(* IEC 61131-3 sources: Industry-PLC-LLM/data/PLCBEAD_repo/PLCBEAD_PLCEmbed-main/PLC-BEAD/Source/PLC_Programs (part 11) *)

(* ---- SIGNAL_4.ST ---- *)
FUNCTION _BYTE_TO_INT:INT
	VAR_INPUT
		IN :	BYTE;
	END_VAR

	_BYTE_TO_INT := USINT_TO_INT(BYTE_TO_USINT(IN));
END_FUNCTION

FUNCTION TIME_TO_UDINT2:UDINT
	VAR_INPUT
		X :	TIME;
	END_VAR

	TIME_TO_UDINT2 := DINT_TO_UDINT(TIME_TO_DINT(X));
END_FUNCTION

FUNCTION UDINT_TO_TIME2:TIME

	VAR_INPUT
		IN :	UDINT;
	END_VAR

	UDINT_TO_TIME2 := DINT_TO_TIME(UDINT_TO_DINT(IN));

END_FUNCTION

FUNCTION_BLOCK T_PLC_MS_block
	VAR_OUTPUT
		T_PLC_MS :	UDINT;
	END_VAR

	VAR_EXTERNAL
		PLC_TICKS_PER_SEC :	INT;
		PLC_SYS_TICK_CNT :	DINT;
	END_VAR

	VAR
		debug :	BOOL;(*Debug-Mode ON / OFF*)
		N :	INT;(*Debug-Faktor*)
		Offset :	UDINT;(*Debug-Offset*)
		temp :	DWORD := DWORD#1;(*Debug-Offset*)
		mode :	BOOL;(*modus*)
		faktor :	UDINT;(*Systemtakt-Faktor*)
		init :	BOOL;
		v_plc_ticks_per_sec :	UDINT;
		base :	UDINT := UDINT#1000;
	END_VAR

	IF init = FALSE THEN
		v_plc_ticks_per_sec := INT_TO_UDINT(PLC_TICKS_PER_SEC);
		IF v_plc_ticks_per_sec = UDINT#1024 THEN
			faktor := UDINT#1;
			mode := FALSE;
		ELSIF v_plc_ticks_per_sec > UDINT#0 THEN
			IF v_plc_ticks_per_sec <= base THEN
				faktor := base / v_plc_ticks_per_sec;
				mode := FALSE;
			ELSE
				faktor := v_plc_ticks_per_sec / base;
				mode := TRUE;
			END_IF;
		ELSE
			faktor := UDINT#1;
		END_IF;
		init := TRUE;
	END_IF;

	IF mode THEN
		T_PLC_MS := DINT_TO_UDINT(PLC_SYS_TICK_CNT) / faktor;
	ELSE
		T_PLC_MS := DINT_TO_UDINT(PLC_SYS_TICK_CNT) * faktor;
	END_IF;

	IF debug THEN
		T_PLC_MS := (DWORD_TO_UDINT(SHL(UDINT_TO_DWORD(T_PLC_MS),N) OR SHL(temp,N)) - UDINT#1) + Offset;
	END_IF;

END_FUNCTION_BLOCK

FUNCTION_BLOCK SIGNAL_Block

	VAR_INPUT
		IN :	BOOL;
		SIG :	BYTE;
		TS :	TIME;
	END_VAR

	VAR_OUTPUT
		Q :	BOOL;
	END_VAR

	VAR
		tx :	DWORD;
		_step :	BYTE;
		T_PLC_MS :	T_PLC_MS_Block;
	END_VAR

	IF in THEN
		T_PLC_MS();
		tx:= UDINT_TO_DWORD(T_PLC_MS.T_PLC_MS);

		IF ts > t#0s THEN
			_step := DWORD_TO_BYTE(UDINT_TO_DWORD(DWORD_TO_UDINT(tx) / TIME_TO_UDINT2(ts)) AND DWORD#16#0000_0007);
		ELSE
			_step := DWORD_TO_BYTE(SHR(tx,7) AND DWORD#16#0000_0007);
		END_IF;
		_step := SHL(BYTE#1,_BYTE_TO_INT(_step));
		Q := (_step AND sig) > BYTE#0;
	ELSE
		Q := FALSE;
	END_IF;

END_FUNCTION_BLOCK

FUNCTION_BLOCK SIGNAL_4_Block

	VAR_INPUT
		IN1 :	BOOL;
		IN2 :	BOOL;
		IN3 :	BOOL;
		IN4 :	BOOL;
		TS :	TIME;
		S1 :	BYTE := 2#1111_1111;
		S2 :	BYTE := 2#1111_0000;
		S3 :	BYTE := 2#1010_1010;
		S4 :	BYTE := 2#1010_0000;
	END_VAR

	VAR_OUTPUT
		Q :	BOOL;
	END_VAR

	VAR
		sig :	SIGNAL_Block;
	END_VAR

	IF in1 THEN
		sig(in := TRUE, sig := s1, TS := TS);
	ELSIF in2 THEN
		sig(in := TRUE, sig := s2, TS := TS);
	ELSIF in3 THEN
		sig(in := TRUE, sig := s3, TS := TS);
	ELSIF in4 THEN
		sig(in := TRUE, sig := s4, TS := TS);
	ELSE
		sig(in := FALSE);
	END_IF;

	Q := sig.Q;

END_FUNCTION_BLOCK

PROGRAM program0

	VAR
		IN1 :	BOOL;
		IN2 :	BOOL;
		IN3 :	BOOL;
		IN4 :	BOOL;
		TS :	TIME;
		S1 :	BYTE := 2#1111_1111;
		S2 :	BYTE := 2#1111_0000;
		S3 :	BYTE := 2#1010_1010;
		S4 :	BYTE := 2#1010_0000;
		Q :	BOOL;
		func_block : SIGNAL_4_Block;
	END_VAR

	func_block.IN1  :=IN1;
	func_block.IN2  :=IN2;
	func_block.IN3  :=IN3;
	func_block.IN4  :=IN4;
	func_block.TS  :=TS;
	func_block.S1  :=S1;
	func_block.S2  :=S2;
	func_block.S3  :=S3;
	func_block.S4  :=S4;
	func_block();
	Q := func_block.Q;

END_PROGRAM

CONFIGURATION Config0

	VAR_GLOBAL
		PLC_TICKS_PER_SEC :	INT;
		PLC_SYS_TICK_CNT :	DINT;
	END_VAR

  	RESOURCE Res0 ON PLC
    	TASK task0(INTERVAL := T#20ms,PRIORITY := 0);
    	PROGRAM instance0 WITH task0 : program0;
  	END_RESOURCE

END_CONFIGURATION

(* ---- SNTP_CLIENT.ST ---- *)
TYPE
  oscat_IP_FIFO128_DATA  : ARRAY [1..128] OF BYTE;
  oscat_Mailbox  : ARRAY [1..16] OF BYTE;

  oscat_IP_FIFO_DATA :
  STRUCT
    X       : oscat_IP_FIFO128_DATA; (* IP_ID FIFO Speicher          *)
    Y       : oscat_IP_FIFO128_DATA; (* IP_ID Z�hler                 *)
    ID      : BYTE;                  (* h�chste vergabene id         *)
    MAX_ID  : BYTE;                  (* maximal Anmeldungen pro ID   *)
      INIT    : BOOL;                  (* Initialisierung durchgef�hrt *)
    EMPTY   : BOOL;                  (* FIFO leer                    *)
    FULL    : BOOL;                  (* FIFO voll                    *)
    TOP     : INT;                   (* maximale anzahl in FIFO      *)
    NW      : INT;                   (* Schreibzeiger                *)
    NR      : INT;                   (* Lesezeiger                   *)
  END_STRUCT;

  oscat_IP_C:
  STRUCT
    C_MODE:			BYTE;          		(*W Mode: TCP/UCP AKTIV/PASSIV                               *)
    C_PORT:         WORD;          		(*W Portnummer                                               *)
    C_IP:           DWORD;         		(*W IP-Adresse gepackt wwxxyyzz = www.xxx.yyy.zzz            *)
    C_STATE:        BYTE;          		(*R Verbindungsstatus ON/OFF + Flanke ON/OFF                 *)
    C_ENABLE:       BOOL;          		(*W Freigabe f�r Connect                                     *)
    R_OBSERVE:      BOOL;          		(*W Empfang ueberwachen                                      *)
    TIME_RESET:     BOOL;          		(*W Alle Timer ruecksetzen                                   *)
    ERROR:          DWORD;         		(*R vvwwxxyy (vv = CON_ERROR, ww = SEN_ERROR, xx = REC_ERROR *)
    FIFO:           oscat_IP_FIFO_DATA; (*I IP FIFO Struktur                                         *)
    MAILBOX:		oscat_Mailbox;		(*I Mailbox: Datenbereich f�r Bausteindatenaustausch         *)
  END_STRUCT;
END_TYPE

TYPE

  oscat_NW_BUF_LONG  : ARRAY [0..4095] OF BYTE;

  oscat_NETWORK_BUFFER :
  STRUCT
    SIZE   : UINT;
    BUFFER : oscat_NW_BUF_LONG;
  END_STRUCT;

END_TYPE

FUNCTION _BYTE_TO_INT:INT
	VAR_INPUT
		IN :	BYTE;
	END_VAR

	_BYTE_TO_INT := USINT_TO_INT(BYTE_TO_USINT(IN));
END_FUNCTION

FUNCTION_BLOCK IP_FIFO_Block

  VAR_IN_OUT
    FIFO :	oscat_IP_FIFO_DATA;
    ID :	BYTE;
    STATE :	BYTE;
  END_VAR

  VAR
    tmp :	INT;
  END_VAR

  IF NOT FIFO.INIT THEN
    FIFO.INIT		:= TRUE;
    FIFO.NW		:= 1;
    FIFO.NR		:= 1;
    FIFO.EMPTY	:= TRUE;
    FIFO.FULL		:= FALSE;
    FIFO.TOP		:= 128;
    FIFO.MAX_ID	:= BYTE#1;
  END_IF;

  IF ID = BYTE#00 THEN
    IF FIFO.ID < INT_TO_BYTE(FIFO.TOP) THEN
      ID := USINT_TO_BYTE(BYTE_TO_USINT(FIFO.ID) + USINT#1);
      FIFO.ID := ID ;

    ELSIF STATE < BYTE#200 THEN
      STATE := BYTE#255;
    RETURN;
    END_IF;
  END_IF;

  IF STATE = BYTE#1 AND NOT FIFO.FULL THEN
    tmp := _BYTE_TO_INT(ID);
    IF FIFO.Y[tmp] < FIFO.MAX_ID THEN
      FIFO.Y[tmp] := USINT_TO_BYTE(BYTE_TO_USINT(FIFO.Y[tmp]) + USINT#1);
      tmp := FIFO.NW;
      FIFO.X[tmp] := ID;
      IF FIFO.NW = FIFO.TOP THEN FIFO.NW := 1; ELSE FIFO.NW := FIFO.NW + 1; END_IF;
      FIFO.FULL := FIFO.NW = FIFO.NR;
    FIFO.EMPTY := FALSE;
      STATE := BYTE#2;
    END_IF;
  END_IF;

  IF STATE = BYTE#2 AND NOT FIFO.EMPTY THEN
    tmp := FIFO.NR;
    IF ID = FIFO.X[tmp] THEN
      STATE := BYTE#3;
    END_IF;
  END_IF;

  IF STATE = BYTE#4 AND NOT FIFO.EMPTY THEN

    tmp := FIFO.NR;
    IF ID = FIFO.X[tmp] THEN
      tmp := _BYTE_TO_INT(ID);
      FIFO.Y[tmp] := USINT_TO_BYTE(BYTE_TO_USINT(FIFO.Y[tmp]) - USINT#1);

      IF FIFO.NR = FIFO.TOP THEN FIFO.NR := 1; ELSE FIFO.NR := FIFO.NR + 1; END_IF;
      FIFO.EMPTY := FIFO.NR = FIFO.NW;
    FIFO.FULL := FALSE;
    END_IF;
    STATE := BYTE#5;
  END_IF;

END_FUNCTION_BLOCK

FUNCTION_BLOCK T_PLC_MS_block

	VAR_OUTPUT
		T_PLC_MS :	UDINT;
	END_VAR

	VAR_EXTERNAL
		PLC_TICKS_PER_SEC :	INT;
		PLC_SYS_TICK_CNT :	DINT;
	END_VAR

	VAR
		debug :	BOOL;(*Debug-Mode ON / OFF*)
		N :	INT;(*Debug-Faktor*)
		Offset :	UDINT;(*Debug-Offset*)
		temp :	DWORD := DWORD#1;(*Debug-Offset*)
		mode :	BOOL;(*modus*)
		faktor :	UDINT;(*Systemtakt-Faktor*)
		init :	BOOL;
		v_plc_ticks_per_sec :	UDINT;
		base :	UDINT := UDINT#1000;
	END_VAR

	IF init = FALSE THEN
		v_plc_ticks_per_sec := INT_TO_UDINT(PLC_TICKS_PER_SEC);
		IF v_plc_ticks_per_sec = UDINT#1024 THEN
			faktor := UDINT#1;
			mode := FALSE;
		ELSIF v_plc_ticks_per_sec > UDINT#0 THEN
			IF v_plc_ticks_per_sec <= base THEN
				faktor := base / v_plc_ticks_per_sec;
				mode := FALSE;
			ELSE
				faktor := v_plc_ticks_per_sec / base;
				mode := TRUE;
			END_IF;
		ELSE
			faktor := UDINT#1;
		END_IF;
		init := TRUE;
	END_IF;

	IF mode THEN
		T_PLC_MS := DINT_TO_UDINT(PLC_SYS_TICK_CNT) / faktor;
	ELSE
		T_PLC_MS := DINT_TO_UDINT(PLC_SYS_TICK_CNT) * faktor;
	END_IF;

	IF debug THEN
		T_PLC_MS := (DWORD_TO_UDINT(SHL(UDINT_TO_DWORD(T_PLC_MS),N) OR SHL(temp,N)) - UDINT#1) + Offset;
	END_IF;

END_FUNCTION_BLOCK

FUNCTION DWORD_OF_BYTE:DWORD
	VAR_INPUT
		B3 :	BYTE;
		B2 :	BYTE;
		B1 :	BYTE;
		B0 :	BYTE;
	END_VAR

	DWORD_OF_BYTE := SHL(SHL(SHL(BYTE_TO_DWORD(B3),8) OR BYTE_TO_DWORD(B2),8) OR BYTE_TO_DWORD(B1),8) OR BYTE_TO_DWORD(B0);

END_FUNCTION

FUNCTION _WORD_TO_DINT:DINT
	VAR_INPUT
		IN :	WORD;
	END_VAR
	_WORD_TO_DINT := UINT_TO_DINT(WORD_TO_UINT(IN));
END_FUNCTION

FUNCTION WORD_OF_BYTE:WORD
	VAR_INPUT
		B1 :	BYTE;
		B0 :	BYTE;
	END_VAR
	WORD_OF_BYTE := SHL(BYTE_TO_WORD(B1),8) OR BYTE_TO_WORD(B0);
END_FUNCTION

FUNCTION _INT_TO_UDINT:UDINT
	VAR_INPUT
		IN :	INT;
	END_VAR

	_INT_TO_UDINT := DINT_TO_UDINT(INT_TO_DINT(IN));
END_FUNCTION

FUNCTION_BLOCK SNTP_CLIENT_Block

  VAR_IN_OUT
    IP_C :	oscat_IP_C;
    S_BUF :	oscat_NETWORK_BUFFER;
    R_BUF :	oscat_NETWORK_BUFFER;
  END_VAR

  VAR_INPUT
    IP4 :	DWORD;
    ACTIVATE :	BOOL;
  END_VAR

  VAR_OUTPUT
    ERROR :	DWORD;
    DONE_P :	BOOL;
    UDT :	UDINT;
    XMS :	INT;
  END_VAR

  VAR
    IP_STATE :	BYTE;
    IP_ID :	BYTE;
    IP_FIFO :	IP_FIFO_Block;
    i :	INT;
    last :	UDINT;
    state :	INT;
    T_PLC_MS :	T_PLC_MS_Block;
    tx :	UDINT;
    ACTIVATE_LAST :	BOOL;
    IP4_STORED :	DWORD;
  END_VAR

  T_PLC_MS();
  tx := T_PLC_MS.T_PLC_MS;

  CASE state OF
  00:
    DONE_P := FALSE;
    IF ACTIVATE AND NOT ACTIVATE_LAST THEN
      IP4_STORED := IP4;
      state := 10;
      ERROR := DWORD#0;
      IP_STATE := BYTE#1;
    END_IF;

  10:
    IF IP_STATE = BYTE#3 THEN

      S_BUF.BUFFER[00] := BYTE#16#1B;
      FOR i := 1 TO 47 DO
        S_BUF.BUFFER[i] := BYTE#16#00;
      END_FOR;

      last := tx;
      state := 30;

      IP_C.C_PORT     := WORD#123;
      IP_C.C_IP       := IP4_STORED;
      IP_C.C_MODE     := BYTE#1;
      IP_C.C_ENABLE   := TRUE;
      IP_C.TIME_RESET := TRUE;
      IP_C.R_OBSERVE  := TRUE;
      S_BUF.SIZE      := UINT#48;
      R_BUF.SIZE      := UINT#0;
    END_IF;

  30:
    IF IP_C.ERROR <> DWORD#00 THEN
      ERROR := IP_C.ERROR;
    S_BUF.SIZE := UINT#0;
    R_BUF.SIZE := UINT#0;
      state := 0;
    ELSIF S_BUF.SIZE = UINT#0 AND R_BUF.SIZE >= UINT#48 THEN
      UDT := DWORD_TO_UDINT(DWORD_OF_BYTE(R_BUF.BUFFER[40],R_BUF.BUFFER[41],R_BUF.BUFFER[42],R_BUF.BUFFER[43]))- UDINT#2208988800;

      XMS := DWORD_TO_INT(SHR(DINT_TO_DWORD(_WORD_TO_DINT(WORD_OF_BYTE(R_BUF.BUFFER[44],R_BUF.BUFFER[45])) * DINT#1000),16));
      XMS := XMS + DWORD_TO_INT(SHR(UDINT_TO_DWORD(tx - last),1));

      UDT := UDT + _INT_TO_UDINT(XMS / 1000);
      XMS := XMS MOD 1000;

      state := 0;
      DONE_P := TRUE;

    END_IF;

    IF state = 0 THEN
      IP_C.R_OBSERVE := FALSE;
      IP_STATE := BYTE#4;
    END_IF;

  END_CASE;

  ACTIVATE_LAST := ACTIVATE;

  IP_FIFO(FIFO:=IP_C.FIFO,STATE:=IP_STATE,ID:=IP_ID);
  IP_C.FIFO:=IP_FIFO.FIFO;
  IP_STATE := IP_FIFO.STATE;
  IP_ID:=IP_FIFO.ID;

END_FUNCTION_BLOCK

PROGRAM program0
	VAR
		IP_C :	oscat_IP_C;
    S_BUF :	oscat_NETWORK_BUFFER;
    R_BUF :	oscat_NETWORK_BUFFER;
    IP4 :	DWORD;
    ACTIVATE :	BOOL;
    ERROR :	DWORD;
    DONE_P :	BOOL;
    UDT :	UDINT;
    XMS :	INT;

		func_block : SNTP_CLIENT_Block;
	END_VAR
	func_block.IP_C := IP_C;
	func_block.S_BUF := S_BUF;
	func_block.R_BUF := R_BUF;
  func_block.IP4 := IP4;
	func_block.ACTIVATE := ACTIVATE;

	func_block();
  IP_C  := func_block.IP_C;
  S_BUF  := func_block.S_BUF;
  R_BUF  := func_block.R_BUF;
  ERROR  := func_block.ERROR;
  DONE_P  := func_block.DONE_P;
  UDT  := func_block.UDT;
  XMS  := func_block.XMS;
END_PROGRAM

CONFIGURATION Config0

	VAR_GLOBAL
		PLC_TICKS_PER_SEC :	INT;
		PLC_SYS_TICK_CNT :	DINT;
	END_VAR

  	RESOURCE Res0 ON PLC
    	TASK task0(INTERVAL := T#20ms,PRIORITY := 0);
    	PROGRAM instance0 WITH task0 : program0;
  	END_RESOURCE

END_CONFIGURATION

(* ---- SNTP_SERVER.ST ---- *)
TYPE
  oscat_IP_FIFO128_DATA  : ARRAY [1..128] OF BYTE;
  oscat_Mailbox  : ARRAY [1..16] OF BYTE;

  oscat_IP_FIFO_DATA :
  STRUCT
    X       : oscat_IP_FIFO128_DATA; (* IP_ID FIFO Speicher          *)
    Y       : oscat_IP_FIFO128_DATA; (* IP_ID Z�hler                 *)
    ID      : BYTE;                  (* h�chste vergabene id         *)
    MAX_ID  : BYTE;                  (* maximal Anmeldungen pro ID   *)
      INIT    : BOOL;                  (* Initialisierung durchgef�hrt *)
    EMPTY   : BOOL;                  (* FIFO leer                    *)
    FULL    : BOOL;                  (* FIFO voll                    *)
    TOP     : INT;                   (* maximale anzahl in FIFO      *)
    NW      : INT;                   (* Schreibzeiger                *)
    NR      : INT;                   (* Lesezeiger                   *)
  END_STRUCT;

  oscat_IP_C:
  STRUCT
    C_MODE:			BYTE;          		(*W Mode: TCP/UCP AKTIV/PASSIV                               *)
    C_PORT:         WORD;          		(*W Portnummer                                               *)
    C_IP:           DWORD;         		(*W IP-Adresse gepackt wwxxyyzz = www.xxx.yyy.zzz            *)
    C_STATE:        BYTE;          		(*R Verbindungsstatus ON/OFF + Flanke ON/OFF                 *)
    C_ENABLE:       BOOL;          		(*W Freigabe f�r Connect                                     *)
    R_OBSERVE:      BOOL;          		(*W Empfang ueberwachen                                      *)
    TIME_RESET:     BOOL;          		(*W Alle Timer ruecksetzen                                   *)
    ERROR:          DWORD;         		(*R vvwwxxyy (vv = CON_ERROR, ww = SEN_ERROR, xx = REC_ERROR *)
    FIFO:           oscat_IP_FIFO_DATA; (*I IP FIFO Struktur                                         *)
    MAILBOX:		oscat_Mailbox;		(*I Mailbox: Datenbereich f�r Bausteindatenaustausch         *)
  END_STRUCT;
END_TYPE

TYPE

  oscat_NW_BUF_LONG  : ARRAY [0..4095] OF BYTE;

  oscat_NETWORK_BUFFER :
  STRUCT
    SIZE   : UINT;
    BUFFER : oscat_NW_BUF_LONG;
  END_STRUCT;

END_TYPE

FUNCTION _BYTE_TO_INT:INT
	VAR_INPUT
		IN :	BYTE;
	END_VAR

	_BYTE_TO_INT := USINT_TO_INT(BYTE_TO_USINT(IN));
END_FUNCTION

FUNCTION_BLOCK IP_FIFO_Block

  VAR_IN_OUT
    FIFO :	oscat_IP_FIFO_DATA;
    ID :	BYTE;
    STATE :	BYTE;
  END_VAR

  VAR
    tmp :	INT;
  END_VAR

  IF NOT FIFO.INIT THEN
    FIFO.INIT		:= TRUE;
    FIFO.NW		:= 1;
    FIFO.NR		:= 1;
    FIFO.EMPTY	:= TRUE;
    FIFO.FULL		:= FALSE;
    FIFO.TOP		:= 128;
    FIFO.MAX_ID	:= BYTE#1;
  END_IF;

  IF ID = BYTE#00 THEN
    IF FIFO.ID < INT_TO_BYTE(FIFO.TOP) THEN
      ID := USINT_TO_BYTE(BYTE_TO_USINT(FIFO.ID) + USINT#1);
      FIFO.ID := ID ;

    ELSIF STATE < BYTE#200 THEN
      STATE := BYTE#255;
    RETURN;
    END_IF;
  END_IF;

  IF STATE = BYTE#1 AND NOT FIFO.FULL THEN
    tmp := _BYTE_TO_INT(ID);
    IF FIFO.Y[tmp] < FIFO.MAX_ID THEN
      FIFO.Y[tmp] := USINT_TO_BYTE(BYTE_TO_USINT(FIFO.Y[tmp]) + USINT#1);
      tmp := FIFO.NW;
      FIFO.X[tmp] := ID;
      IF FIFO.NW = FIFO.TOP THEN FIFO.NW := 1; ELSE FIFO.NW := FIFO.NW + 1; END_IF;
      FIFO.FULL := FIFO.NW = FIFO.NR;
    FIFO.EMPTY := FALSE;
      STATE := BYTE#2;
    END_IF;
  END_IF;

  IF STATE = BYTE#2 AND NOT FIFO.EMPTY THEN
    tmp := FIFO.NR;
    IF ID = FIFO.X[tmp] THEN
      STATE := BYTE#3;
    END_IF;
  END_IF;

  IF STATE = BYTE#4 AND NOT FIFO.EMPTY THEN

    tmp := FIFO.NR;
    IF ID = FIFO.X[tmp] THEN
      tmp := _BYTE_TO_INT(ID);
      FIFO.Y[tmp] := USINT_TO_BYTE(BYTE_TO_USINT(FIFO.Y[tmp]) - USINT#1);

      IF FIFO.NR = FIFO.TOP THEN FIFO.NR := 1; ELSE FIFO.NR := FIFO.NR + 1; END_IF;
      FIFO.EMPTY := FIFO.NR = FIFO.NW;
    FIFO.FULL := FALSE;
    END_IF;
    STATE := BYTE#5;
  END_IF;

END_FUNCTION_BLOCK

FUNCTION_BLOCK T_PLC_MS_block

	VAR_OUTPUT
		T_PLC_MS :	UDINT;
	END_VAR

	VAR_EXTERNAL
		PLC_TICKS_PER_SEC :	INT;
		PLC_SYS_TICK_CNT :	DINT;
	END_VAR

	VAR
		debug :	BOOL;(*Debug-Mode ON / OFF*)
		N :	INT;(*Debug-Faktor*)
		Offset :	UDINT;(*Debug-Offset*)
		temp :	DWORD := DWORD#1;(*Debug-Offset*)
		mode :	BOOL;(*modus*)
		faktor :	UDINT;(*Systemtakt-Faktor*)
		init :	BOOL;
		v_plc_ticks_per_sec :	UDINT;
		base :	UDINT := UDINT#1000;
	END_VAR

	IF init = FALSE THEN
		v_plc_ticks_per_sec := INT_TO_UDINT(PLC_TICKS_PER_SEC);
		IF v_plc_ticks_per_sec = UDINT#1024 THEN
			faktor := UDINT#1;
			mode := FALSE;
		ELSIF v_plc_ticks_per_sec > UDINT#0 THEN
			IF v_plc_ticks_per_sec <= base THEN
				faktor := base / v_plc_ticks_per_sec;
				mode := FALSE;
			ELSE
				faktor := v_plc_ticks_per_sec / base;
				mode := TRUE;
			END_IF;
		ELSE
			faktor := UDINT#1;
		END_IF;
		init := TRUE;
	END_IF;

	IF mode THEN
		T_PLC_MS := DINT_TO_UDINT(PLC_SYS_TICK_CNT) / faktor;
	ELSE
		T_PLC_MS := DINT_TO_UDINT(PLC_SYS_TICK_CNT) * faktor;
	END_IF;

	IF debug THEN
		T_PLC_MS := (DWORD_TO_UDINT(SHL(UDINT_TO_DWORD(T_PLC_MS),N) OR SHL(temp,N)) - UDINT#1) + Offset;
	END_IF;

END_FUNCTION_BLOCK

FUNCTION_BLOCK SNTP_SERVER_Block

  VAR_IN_OUT
    IP_C :	oscat_IP_C;
    S_BUF :	oscat_NETWORK_BUFFER;
    R_BUF :	oscat_NETWORK_BUFFER;
  END_VAR

  VAR_INPUT
    ENABLE :	BOOL;
    STRATUM :	BYTE := BYTE#1;
    UDT :	UDINT;
    XMS :	INT;
  END_VAR

  VAR
    IP_STATE :	BYTE;
    IP_ID :	BYTE;
    IP_FIFO :	IP_FIFO_Block;
    i2 :	INT;
    i :	INT;
    TIMESTAMP_INT :	DWORD;
    TIMESTAMP_SEK :	DWORD;
    TS_B :	BYTE;
    state :	INT;
    T_PLC_MS :	T_PLC_MS_Block;
    tx :	UDINT;
    t :	TON;
  END_VAR

  T_PLC_MS();
  tx := T_PLC_MS.T_PLC_MS;

  CASE state OF

  00:
    IF ENABLE THEN
      state := 10;
      IP_STATE := BYTE#1;
    END_IF;

  10:
    IF IP_STATE = BYTE#3 THEN

      IP_C.C_PORT     := WORD#123;
      IP_C.C_IP       := DWORD#00;
      IP_C.C_MODE     := BYTE#5;
      IP_C.C_ENABLE   := TRUE;
      IP_C.TIME_RESET := TRUE;
      IP_C.R_OBSERVE  := FALSE;
      S_BUF.SIZE      := UINT#0;
      R_BUF.SIZE      := UINT#0;

      state := 20;
    END_IF;

  20:
    IF R_BUF.SIZE > UINT#0 THEN
      state := 20;
      FOR i := 0 TO 47 DO
        IF INT_TO_UINT(i) > R_BUF.SIZE - UINT#1 THEN
          R_BUF.BUFFER[i] := BYTE#00;
      END_IF;
        S_BUF.BUFFER[i] := BYTE#00;
      END_FOR;

    R_BUF.SIZE := UINT#0;

      S_BUF.BUFFER[0] := BYTE#2#11100;
      S_BUF.BUFFER[1] := STRATUM;
      S_BUF.BUFFER[2] := BYTE#10;
      S_BUF.BUFFER[3] := BYTE#16#FB;

      TIMESTAMP_INT := UDINT_TO_DWORD(UDT + UDINT#2208988800);

    TIMESTAMP_SEK := DINT_TO_DWORD(DWORD_TO_DINT(SHL(INT_TO_DWORD(XMS),16))/DINT#1000);

      TS_B := TIMESTAMP_INT.B3;
      S_BUF.BUFFER[16] := TS_B;
      S_BUF.BUFFER[32] := TS_B;
      S_BUF.BUFFER[40] := TS_B;

      TS_B := TIMESTAMP_INT.B2;
      S_BUF.BUFFER[17] := TS_B;
      S_BUF.BUFFER[33] := TS_B;
      S_BUF.BUFFER[41] := TS_B;

      TS_B := TIMESTAMP_INT.B1;
      S_BUF.BUFFER[18] := TS_B;
      S_BUF.BUFFER[34] := TS_B;
      S_BUF.BUFFER[42] := TS_B;

      TS_B := TIMESTAMP_INT.B0;
      S_BUF.BUFFER[19] := TS_B;
      S_BUF.BUFFER[35] := TS_B;
      S_BUF.BUFFER[43] := TS_B;

      TS_B := TIMESTAMP_SEK.B1;
      S_BUF.BUFFER[20] := TS_B;
      S_BUF.BUFFER[36] := TS_B;
      S_BUF.BUFFER[44] := TS_B;

      TS_B := TIMESTAMP_SEK.B0;
      S_BUF.BUFFER[21] := TS_B;
      S_BUF.BUFFER[37] := TS_B;
      S_BUF.BUFFER[45] := TS_B;

      i2 := 40;
      FOR i := 24 TO 31 DO
        S_BUF.BUFFER[i] := R_BUF.BUFFER[i2];
        i2 := i2 +1;
      END_FOR;

      S_BUF.SIZE := UINT#48;

    ELSIF NOT ENABLE AND S_BUF.SIZE = UINT#0 THEN
      IP_STATE := BYTE#4;
      state := 0;
    END_IF;

  END_CASE;

  t(IN:= IP_C.ERROR > DWORD#0, PT:=T#5s);
  IF t.Q THEN
    IP_C.TIME_RESET := TRUE;
  END_IF;

  IP_FIFO(FIFO:=IP_C.FIFO,STATE:=IP_STATE,ID:=IP_ID);
  IP_C.FIFO:=IP_FIFO.FIFO;
  IP_STATE := IP_FIFO.STATE;
  IP_ID:=IP_FIFO.ID;

END_FUNCTION_BLOCK

PROGRAM program0
	VAR
		IP_C :	oscat_IP_C;
    S_BUF :	oscat_NETWORK_BUFFER;
    R_BUF :	oscat_NETWORK_BUFFER;
    ENABLE :	BOOL;
    STRATUM :	BYTE := BYTE#1;
    UDT :	UDINT;
    XMS :	INT;

		func_block : SNTP_SERVER_Block;
	END_VAR
	func_block.IP_C := IP_C;
	func_block.S_BUF := S_BUF;
	func_block.R_BUF := R_BUF;
  func_block.ENABLE := ENABLE;
	func_block.STRATUM := STRATUM;
	func_block.UDT := UDT;
  func_block.XMS := XMS;

	func_block();
  IP_C  := func_block.IP_C;
  S_BUF  := func_block.S_BUF;
  R_BUF  := func_block.R_BUF;
END_PROGRAM

CONFIGURATION Config0

	VAR_GLOBAL
		PLC_TICKS_PER_SEC :	INT;
		PLC_SYS_TICK_CNT :	DINT;
	END_VAR

  	RESOURCE Res0 ON PLC
    	TASK task0(INTERVAL := T#20ms,PRIORITY := 0);
    	PROGRAM instance0 WITH task0 : program0;
  	END_RESOURCE

END_CONFIGURATION

(* ---- SPEED.ST ---- *)
FUNCTION_BLOCK SPEED_Block

	VAR_INPUT
		MS :	REAL;
		KMH :	REAL;
		KN :	REAL;
		MH :	REAL;
	END_VAR

	VAR_OUTPUT
		YMS :	REAL;
		YKMH :	REAL;
		YKN :	REAL;
		YMH :	REAL;
	END_VAR

	Yms := ms +
			kmh * 0.27777777777778 +
			kn * 0.5144444 +
			mh * 0.44704;
	Ykmh := Yms * 3.6;
	Ykn := Yms * 1.94384466037535;
	Ymh := Yms * 2.23693629205440;

END_FUNCTION_BLOCK

PROGRAM program0

	VAR
		MS :	REAL;
		KMH :	REAL;
		KN :	REAL;
		MH :	REAL;
		YMS :	REAL;
		YKMH :	REAL;
		YKN :	REAL;
		YMH :	REAL;
		func_block : SPEED_Block;
	END_VAR
		func_block.MS  :=MS;
		func_block.KMH  :=KMH;
		func_block.KN  :=KN;
		func_block.MH  :=MH;
		func_block();
		YMS := func_block.YMS;
		YKMH := func_block.YKMH;
		YKN := func_block.YKN;
		YMH := func_block.YMH;

	END_PROGRAM

CONFIGURATION Config0

	RESOURCE Res0 ON PLC
		TASK task0(INTERVAL := T#20ms,PRIORITY := 0);
		PROGRAM instance0 WITH task0 : program0;
	END_RESOURCE

END_CONFIGURATION

(* ---- SRAMP.ST ---- *)
FUNCTION_BLOCK T_PLC_US_Block
	VAR_OUTPUT
		T_PLC_US :	UDINT;
	END_VAR

	VAR_EXTERNAL
		PLC_TICKS_PER_SEC :	INT;
		PLC_SYS_TICK_CNT :	DINT;
	END_VAR

	VAR
		debug :	BOOL;
		N :	INT;
		Offset :	UDINT;
		temp :	DWORD := DWORD#1;
		mode :	BOOL;
		faktor :	UDINT;
		init :	BOOL;
		v_plc_ticks_per_sec :	UDINT;
		base :	UDINT := UDINT#1000000;
	END_VAR

	IF init = FALSE THEN
		v_plc_ticks_per_sec := INT_TO_UDINT(PLC_TICKS_PER_SEC);
		IF v_plc_ticks_per_sec = UDINT#1024 THEN
			faktor := UDINT#1000;
			mode := FALSE;
		ELSIF v_plc_ticks_per_sec > UDINT#0 THEN
			IF v_plc_ticks_per_sec <= base THEN
				faktor := base / v_plc_ticks_per_sec;
				mode := FALSE;
			ELSE
				faktor := v_plc_ticks_per_sec / base;
				mode := TRUE;
			END_IF;
		ELSE
			faktor := UDINT#1;
		END_IF;
		init := TRUE;
	END_IF;

	IF mode THEN
		T_PLC_US := DINT_TO_UDINT(PLC_SYS_TICK_CNT) / faktor;
	ELSE
		T_PLC_US := DINT_TO_UDINT(PLC_SYS_TICK_CNT) * faktor;
	END_IF;

	IF debug THEN
		T_PLC_US := (DWORD_TO_UDINT(SHL(UDINT_TO_DWORD(T_PLC_US),N) OR SHL(temp,N)) - UDINT#1) + Offset;
	END_IF;
END_FUNCTION_BLOCK

FUNCTION_BLOCK TC_S_Block

	VAR_OUTPUT
		TC :	REAL;
	END_VAR

	VAR
		init :	BOOL;
		tx :	UDINT;
		last :	UDINT;
		T_PLC_US :	T_PLC_US_Block;
	END_VAR

	T_PLC_US();
	tx:= T_PLC_US.T_PLC_US;

	IF NOT init THEN
		init := TRUE;
		TC := 0.0;
	ELSE
		tc := UDINT_TO_REAL(tx - last) * 1.0E-6;
	END_IF;
	last := tx;

END_FUNCTION_BLOCK

FUNCTION_BLOCK SRAMP_Block

	VAR_INPUT
		X :	REAL;
		A_UP :	REAL;
		A_DN :	REAL;
		VU_MAX :	REAL;
		VD_MAX :	REAL;
		LIMIT_HIGH :	REAL;
		LIMIT_LOW :	REAL;
		RST :	BOOL;
	END_VAR

	VAR_OUTPUT
		Y :	REAL;
		V :	REAL;
	END_VAR

	VAR
		cycle_time :	TC_S_Block;
		init :	BOOL;
	END_VAR

	cycle_time();

	A_up := MAX(0.0,A_UP);
	A_dn := MIN(0.0,A_dn);
	VU_max := MAX(0.0,VU_max);
	VD_max := MIN(0.0,VD_MAX);

	IF rst OR NOT init THEN
		init := TRUE;
		Y := 0.0;
		V := 0.0;
	ELSIF X = Y THEN
		v := 0.0;
	ELSIF X > Y THEN
		v := MIN(v + A_UP * cycle_time.TC, vu_max);
		v := MIN(SQRT((Y-X) * 2.0 * A_DN), v);
		y := LIMIT(limit_low, y + MIN(v * cycle_time.TC, X-Y), limit_high);
	ELSIF X < Y THEN
		v := MAX(v + A_DN * cycle_time.TC, vd_max);
		v := MAX(-SQRT((Y-X) * 2.0 * A_UP), v);
		y := LIMIT(limit_low, y + MAX(v * cycle_time.TC, X-Y), limit_high);
	END_IF;

END_FUNCTION_BLOCK

PROGRAM program0
	VAR
		X :	REAL;
		A_UP :	REAL;
		A_DN :	REAL;
		VU_MAX :	REAL;
		VD_MAX :	REAL;
		LIMIT_HIGH :	REAL;
		LIMIT_LOW :	REAL;
		RST :	BOOL;
		Y :	REAL;
		V :	REAL;
		func_block : SRAMP_Block;
	END_VAR
		func_block.X  := X;
		func_block.A_UP  := A_UP;
		func_block.A_DN  := A_DN;
		func_block.VU_MAX  := VU_MAX;
		func_block.VD_MAX  := VD_MAX;
		func_block.LIMIT_HIGH  := LIMIT_HIGH;
		func_block.LIMIT_LOW  := LIMIT_LOW;
		func_block.RST  := RST;
		func_block();
		Y := func_block.Y;
		V := func_block.V;

END_PROGRAM

CONFIGURATION Config0

	VAR_GLOBAL
		PLC_TICKS_PER_SEC :	INT;
		PLC_SYS_TICK_CNT :	DINT;
	END_VAR

	RESOURCE Res0 ON PLC
		TASK task0(INTERVAL := T#20ms,PRIORITY := 0);
		PROGRAM instance0 WITH task0 : program0;
	END_RESOURCE

END_CONFIGURATION

(* ---- STACK_16.ST ---- *)
TYPE
  oscat_ardw_0_15             : ARRAY [0..15]   OF DWORD;
END_TYPE

FUNCTION_BLOCK STACK_16_Block

	VAR_INPUT
		DIN :	DWORD;
		E :	BOOL := TRUE;
		RD :	BOOL;
		WD :	BOOL;
		RST :	BOOL;
	END_VAR

	VAR_OUTPUT
		DOUT :	DWORD;
		EMPTY :	BOOL := TRUE;
		FULL :	BOOL;
	END_VAR

	VAR
		pt :	INT;
		stack :	oscat_ardw_0_15;
	END_VAR

	IF RST THEN
		pt := 0;
		EMPTY := TRUE;
		FULL := FALSE;
		Dout := DWORD#0;
	ELSIF E THEN
		IF NOT EMPTY AND RD THEN
			pt := pt - 1;
			Dout := stack[pt];
			EMPTY := pt = 0;
			FULL := FALSE;
		END_IF;
		IF NOT FULL AND WD THEN
			stack[pt] := Din;
			pt := pt + 1;
			FULL := pt > 15;
			EMPTY := FALSE;
		END_IF;
	END_IF;

END_FUNCTION_BLOCK

PROGRAM program0
	VAR
		DIN :	DWORD;
		E :	BOOL := TRUE;
		RD :	BOOL;
		WD :	BOOL;
		RST :	BOOL;
		DOUT :	DWORD;
		EMPTY :	BOOL := TRUE;
		FULL :	BOOL;
		func_block : STACK_16_Block;
	END_VAR
		func_block.DIN  := DIN;
		func_block.E  := E;
		func_block.RD  := RD;
		func_block.WD  := WD;
		func_block.RST  := RST;
		func_block();
		DOUT := func_block.DOUT;
		EMPTY := func_block.EMPTY;
		FULL := func_block.FULL;

END_PROGRAM

CONFIGURATION Config0

	RESOURCE Res0 ON PLC
		TASK task0(INTERVAL := T#20ms,PRIORITY := 0);
		PROGRAM instance0 WITH task0 : program0;
	END_RESOURCE

END_CONFIGURATION

(* ---- STACK_32.ST ---- *)
TYPE
  	oscat_ardw_0_31             : ARRAY [0..31]   OF DWORD;
END_TYPE

FUNCTION_BLOCK STACK_32_Block

	VAR_INPUT
		DIN :	DWORD;
		E :	BOOL := TRUE;
		RD :	BOOL;
		WD :	BOOL;
		RST :	BOOL;
	END_VAR

	VAR_OUTPUT
		DOUT :	DWORD;
		EMPTY :	BOOL := TRUE;
		FULL :	BOOL;
	END_VAR

	VAR
		pt :	INT;
		stack :	oscat_ardw_0_31;
	END_VAR

	IF RST THEN
		pt := 0;
		EMPTY := TRUE;
		FULL := FALSE;
		Dout := DWORD#0;
	ELSIF E THEN
		IF NOT EMPTY AND RD THEN
			(* read one element *)
			pt := pt - 1;
			Dout := stack[pt];
			EMPTY := pt = 0;
			FULL := FALSE;
		END_IF;
		IF NOT FULL AND WD THEN
			(* write one element *)
			stack[pt] := Din;
			pt := pt + 1;
			FULL := pt > 31;
			EMPTY := FALSE;
		END_IF;
	END_IF;

END_FUNCTION_BLOCK

PROGRAM program0
	VAR
		DIN :	DWORD;
		E :	BOOL := TRUE;
		RD :	BOOL;
		WD :	BOOL;
		RST :	BOOL;
		DOUT :	DWORD;
		EMPTY :	BOOL := TRUE;
		FULL :	BOOL;
		func_block : STACK_32_Block;
	END_VAR
		func_block.DIN  := DIN;
		func_block.E  := E;
		func_block.RD  := RD;
		func_block.WD  := WD;
		func_block.RST  := RST;
		func_block();
		DOUT := func_block.DOUT;
		EMPTY := func_block.EMPTY;
		FULL := func_block.FULL;

END_PROGRAM

CONFIGURATION Config0

	RESOURCE Res0 ON PLC
		TASK task0(INTERVAL := T#20ms,PRIORITY := 0);
		PROGRAM instance0 WITH task0 : program0;
	END_RESOURCE

END_CONFIGURATION

(* ---- STAIR2.ST ---- *)
FUNCTION FLOOR : INT
	VAR_INPUT
		x : REAL;
	END_VAR

	FLOOR := REAL_TO_INT(X);
	IF INT_TO_REAL(FLOOR) > X THEN
		floor := floor - 1;
	END_IF;
END_FUNCTION

FUNCTION_BLOCK STAIR2_Block

	VAR_INPUT
		X :	REAL;
		D :	REAL;
	END_VAR

	VAR_OUTPUT
		Y :	REAL;
	END_VAR

	IF D > 0.0 THEN
		IF X >= Y + D OR X <= Y - D THEN Y := INT_TO_REAL(FLOOR(X/D)) * D; END_IF;
	ELSE
		Y := X;
	END_IF;

END_FUNCTION_BLOCK

PROGRAM program0

	VAR
		X :	REAL;
		D :	REAL;
		Y :	REAL;
		func_block : STAIR2_Block;
	END_VAR
	func_block.X := X;
	func_block.D := D;
	func_block();
	Y := func_block.Y;

END_PROGRAM

CONFIGURATION Config0

	RESOURCE Res0 ON PLC
		TASK task0(INTERVAL := T#20ms,PRIORITY := 0);
		PROGRAM instance0 WITH task0 : program0;
	END_RESOURCE

END_CONFIGURATION

(* ---- STATUS_TO_ESR.ST ---- *)
TYPE
  oscat_esr_collect_data      : ARRAY [0..7]    OF BYTE;
END_TYPE

TYPE oscat_esr_data :
  STRUCT
	typ    : BYTE;
	adress : STRING;
	DS     : UDINT;
	TS     : TIME;
	data   : oscat_esr_collect_data;
  END_STRUCT;
END_TYPE

FUNCTION_BLOCK STATUS_TO_ESR_Block

	VAR_INPUT
		STATUS :	BYTE;
		ADRESS :	STRING;
		DT_IN :	UDINT;
		TS :	TIME;
	END_VAR

	VAR_OUTPUT
		STATUS_TO_ESR :	oscat_esr_data;
	END_VAR

	IF status < BYTE#100 THEN
		status_to_ESR.typ := BYTE#1;
	ELSIF status < BYTE#200 THEN
		status_to_ESR.typ := BYTE#2;
	ELSE
		status_to_ESR.typ := BYTE#3;
	END_IF;
	status_to_ESR.adress:= adress;
	status_to_ESR.DS := DT_in;
	status_to_ESR.TS := TS;
	status_to_ESR.data[0] := status;
END_FUNCTION_BLOCK

PROGRAM program0
	VAR
		STATUS :	BYTE;
		ADRESS :	STRING;
		DT_IN  :	UDINT;
		TS     :	TIME;
		STATUS_TO_ESR :	oscat_esr_data;

		func_block : STATUS_TO_ESR_Block;
	END_VAR
	func_block.STATUS := STATUS;
	func_block.ADRESS := ADRESS;
	func_block.DT_IN := DT_IN ;
	func_block.TS    := TS    ;

	func_block();
	STATUS_TO_ESR  := func_block.STATUS_TO_ESR;
END_PROGRAM

CONFIGURATION Config0
	RESOURCE Res0 ON PLC
		TASK task0(INTERVAL := T#20ms,PRIORITY := 0);
		PROGRAM instance0 WITH task0 : program0;
	END_RESOURCE
END_CONFIGURATION

(* ---- STORE_8.ST ---- *)
FUNCTION_BLOCK STORE_8_Block

	VAR_INPUT
		SET :	BOOL;
		D0 :	BOOL;
		D1 :	BOOL;
		D2 :	BOOL;
		D3 :	BOOL;
		D4 :	BOOL;
		D5 :	BOOL;
		D6 :	BOOL;
		D7 :	BOOL;
		CLR :	BOOL;
		RST :	BOOL;
	END_VAR

	VAR_OUTPUT
		Q0 :	BOOL;
		Q1 :	BOOL;
		Q2 :	BOOL;
		Q3 :	BOOL;
		Q4 :	BOOL;
		Q5 :	BOOL;
		Q6 :	BOOL;
		Q7 :	BOOL;
	END_VAR

	VAR
		edge :	BOOL;
	END_VAR

	IF rst OR set THEN
		q0 := NOT rst;
		q1 := q0;
		q2 := q0;
		q3 := q0;
		q4 := q0;
		q5 := q0;
		q6 := q0;
		q7 := q0;
	ELSE
		IF D0 THEN Q0 := TRUE; END_IF;
		IF D1 THEN Q1 := TRUE; END_IF;
		IF D2 THEN Q2 := TRUE; END_IF;
		IF D3 THEN Q3 := TRUE; END_IF;
		IF D4 THEN Q4 := TRUE; END_IF;
		IF D5 THEN Q5 := TRUE; END_IF;
		IF D6 THEN Q6 := TRUE; END_IF;
		IF D7 THEN Q7 := TRUE; END_IF;

		IF clr AND NOT edge THEN
			IF q0 THEN q0 := FALSE;
			ELSIF q1 THEN q1 := FALSE;
			ELSIF q2 THEN q2 := FALSE;
			ELSIF q3 THEN q3 := FALSE;
			ELSIF q4 THEN q4 := FALSE;
			ELSIF q5 THEN q5 := FALSE;
			ELSIF q6 THEN q6 := FALSE;
			ELSE q7 := FALSE;
			END_IF;
		END_IF;
		edge := clr;
	END_IF;

END_FUNCTION_BLOCK

PROGRAM program0
	VAR
		SET :	BOOL;
		D0 :	BOOL;
		D1 :	BOOL;
		D2 :	BOOL;
		D3 :	BOOL;
		D4 :	BOOL;
		D5 :	BOOL;
		D6 :	BOOL;
		D7 :	BOOL;
		CLR :	BOOL;
		RST :	BOOL;
		Q0 :	BOOL;
		Q1 :	BOOL;
		Q2 :	BOOL;
		Q3 :	BOOL;
		Q4 :	BOOL;
		Q5 :	BOOL;
		Q6 :	BOOL;
		Q7 :	BOOL;
		func_block : STORE_8_Block;
	END_VAR
	func_block.SET  := SET;
	func_block.D0  := D0;
	func_block.D1  := D1;
	func_block.D2  := D2;
	func_block.D3  := D3;
	func_block.D4  := D4;
	func_block.D5  := D5;
	func_block.D6  := D6;
	func_block.D7  := D7;
	func_block.CLR  := CLR;
	func_block.RST  := RST;
	func_block();
	Q0  := func_block.Q0;
	Q1  := func_block.Q1;
	Q2  := func_block.Q2;
	Q3  := func_block.Q3;
	Q4  := func_block.Q4;
	Q5  := func_block.Q5;
	Q6  := func_block.Q6;
	Q7  := func_block.Q7;
END_PROGRAM

CONFIGURATION Config0
	RESOURCE Res0 ON PLC
		TASK task0(INTERVAL := T#20ms,PRIORITY := 0);
		PROGRAM instance0 WITH task0 : program0;
	END_RESOURCE
END_CONFIGURATION

(* ---- STRING_TO_BUFFER.ST ---- *)
TYPE
	oscat_STRING250             : STRING(250);
	oscat_arb_0_249 			  : ARRAY [0..249] 	OF BYTE;
END_TYPE

FUNCTION_BLOCK _STRING_TO_BUFFER_Block
	VAR_INPUT
		STR :	oscat_STRING250;
		POS :	INT;
		SIZE :	UINT;
	END_VAR

	VAR_OUTPUT
		_STRING_TO_BUFFER :	INT;
	END_VAR

	VAR_IN_OUT
		PT :	oscat_arb_0_249;
	END_VAR

	VAR
		i :	INT;
		end :	INT;
		x :	INT;
	END_VAR

	IF pos < 0 THEN RETURN; END_IF;
	end := MIN(pos + LEN(str), UINT_TO_INT(size)) - 1;
	x:= 1;
	FOR i := pos TO end DO
		pt[i] := INT_TO_BYTE(GET_CHAR(str,x));
		x := x + 1;
	END_FOR;

	_STRING_TO_BUFFER := i;
END_FUNCTION_BLOCK

PROGRAM program0
	VAR
	    LocalVar1 : oscat_STRING250;
        LocalVar2 : INT;
        LocalVar3 : UINT;
		LocalInOut : oscat_arb_0_249;
		LocalOUT  : INT;
		func_block : _STRING_TO_BUFFER_Block;
  	END_VAR
	func_block.STR := LocalVar1;
    func_block.POS := LocalVar2;
    func_block.SIZE := LocalVar3;
	func_block.PT := LocalInOut;
	func_block();
	LocalOUT := func_block._STRING_TO_BUFFER;
	LocalInOut := func_block.PT;
END_PROGRAM

CONFIGURATION Config0
  	RESOURCE Res0 ON PLC
    	TASK task0(INTERVAL := T#20ms,PRIORITY := 0);
    	PROGRAM instance0 WITH task0 : program0;
  	END_RESOURCE
END_CONFIGURATION

(* ---- STRING_TO_TIME.ST ---- *)
FUNCTION_BLOCK UPPERCASE_Block

	VAR_INPUT
		STR :	STRING;
	END_VAR

	VAR_OUTPUT
		UPPERCASE :	STRING;
	END_VAR

	VAR
		char :	BYTE;
		char2 :	BYTE;
		pos :	INT;
		l :	INT;
		str_temp :	STRING;
	END_VAR

	UPPERCASE := str;
	l := LEN(str);
	FOR pos := 1 TO l DO
		char := INT_TO_BYTE(GET_CHAR(str,pos));
		char2 := TO_UPPER(char);
		IF char <> char2 THEN
			str_temp := UPPERCASE;
			UPPERCASE := REPLACE(str_temp,BYTE_TO_STRING(char2,'%c'),1,pos);
		END_IF;
	END_FOR;

END_FUNCTION_BLOCK

FUNCTION_BLOCK _STRING_TO_TIME
  VAR_INPUT
    _TIME :	STRING;
  END_VAR

  VAR_OUTPUT
    STRING_TO_TIME_O :	TIME;
  END_VAR

  VAR
    pos1 :	INT;
    pos2 :	INT;
    tmp :	STRING;
    tmp2 :	STRING;
    UPPERCASE :	UPPERCASE_Block;
    FINDB_NONUM :	FINDB_NONUM;
    FINDB_NUM :	FINDB_NUM;
    faktor :	UDINT;
    IS_ALNUM :	IS_ALNUM;
  END_VAR

  UPPERCASE(str:=_TIME);
  tmp:=UPPERCASE.UPPERCASE;

  STRING_TO_TIME_O := T#0s;

  WHILE (TRUE) DO
    FAKTOR := UDINT#0;

    FINDB_NONUM(str:=tmp);
    pos2:=FINDB_NONUM.findB_nonum;

    FINDB_NUM(str:=tmp);
    pos1:=FINDB_NUM.findB_num;

    (* bezeichner gefunden *)
    IF POS1>0 AND (POS2>POS1) THEN

      tmp2 := RIGHT(tmp,POS2-POS1);
      tmp := LEFT(tmp,pos1);

      IF EQ_STRING(tmp2,'MS') THEN
      FAKTOR := UDINT#1;
      ELSIF EQ_STRING(tmp2,'S') THEN
      FAKTOR := UDINT#1000;
      ELSIF EQ_STRING(tmp2,'M') THEN
      FAKTOR := UDINT#60000;
      ELSIF EQ_STRING(tmp2,'H') THEN
      FAKTOR := UDINT#3600000;
      ELSIF EQ_STRING(tmp2,'D') THEN
      FAKTOR := UDINT#864000000;
      END_IF;
    ELSE
      EXIT;
    END_IF;

    IF FAKTOR > UDINT#0 THEN

      FINDB_NONUM(str:=tmp);
      pos1:=FINDB_NONUM.findB_nonum;
      IF pos1>0 THEN
        tmp2 := RIGHT(tmp,LEN(tmp)-pos1);
        tmp := LEFT(tmp,pos1);
        IS_ALNUM(str:=tmp2);
        IF IS_ALNUM.IS_ALNUM THEN
          STRING_TO_TIME_O := STRING_TO_TIME_O + UDINT_TO_TIME(faktor * STRING_TO_UDINT(tmp2));
        END_IF;
      ELSE
      EXIT;
      END_IF;
    END_IF;
  END_WHILE;
END_FUNCTION_BLOCK

PROGRAM program0
	VAR
    LocalVar1 : STRING;
		LocalOUT  : TIME;
		func_block : _INSERT80;
  	END_VAR
	func_block._TIME := LocalVar1;
	func_block();
	LocalOUT := func_block.STRING_TO_TIME_O;
END_PROGRAM

CONFIGURATION Config0
  	RESOURCE Res0 ON PLC
    	TASK task0(INTERVAL := T#20ms,PRIORITY := 0);
    	PROGRAM instance0 WITH task0 : program0;
  	END_RESOURCE
END_CONFIGURATION

(* ---- STRING_TO_TOD.ST ---- *)
FUNCTION_BLOCK STRING_TO_TOD_Block

  VAR_INPUT
    _TOD :	STRING;
  END_VAR

  VAR_OUTPUT
    out_STRING_TO_TOD :	UDINT;
  END_VAR

  VAR
    pos :	INT;
    i :	INT;
    tmp :	STRING;
    tmp2 :	STRING;
  END_VAR

  out_STRING_TO_TOD := UDINT#0;
  i := LEN(_TOD);
  pos :=FIND(_TOD,'#');

  IF pos>0 AND i>pos THEN
    tmp := RIGHT(_TOD,LEN(_TOD)-pos);
    pos := FIND(tmp,':');
    IF pos>1 THEN
      tmp2 := LEFT(tmp,pos-1);
      tmp := RIGHT(tmp,LEN(tmp)-pos);
      out_STRING_TO_TOD := STRING_TO_UDINT(tmp2) * UDINT#3600000;

      pos :=FIND(tmp,':');
      IF pos>1 THEN
        tmp2 := LEFT(tmp,pos-1);
        tmp := RIGHT(tmp,LEN(tmp)-pos);
        out_STRING_TO_TOD := out_STRING_TO_TOD + STRING_TO_UDINT(tmp2) * UDINT#60000;

        out_STRING_TO_TOD := out_STRING_TO_TOD + STRING_TO_UDINT(tmp) * UDINT#1000;
      END_IF;
    END_IF;
  END_IF;

END_FUNCTION_BLOCK

PROGRAM program0
  VAR
    _TOD :	STRING;
  	out_STRING_TO_TOD :	UDINT;
    func_block : STRING_TO_TOD_Block;
  END_VAR
	func_block._TOD  := _TOD;
	func_block();
	out_STRING_TO_TOD  := func_block.out_STRING_TO_TOD;
END_PROGRAM

CONFIGURATION Config0
	RESOURCE Res0 ON PLC
		TASK task0(INTERVAL := T#20ms,PRIORITY := 0);
		PROGRAM instance0 WITH task0 : program0;
	END_RESOURCE
END_CONFIGURATION

(* ---- STRING_TO_URL.ST ---- *)
TYPE
  oscat_STRING250             : STRING;
  oscat_STRING32             : STRING;
  oscat_STRING80             : STRING;
  oscat_STRING160             : STRING;
  oscat_STRING40             : STRING;
  oscat_STRING10             : STRING;
  oscat_STRING20             : STRING;
END_TYPE

TYPE oscat_url :
    STRUCT
    PROTOCOL : oscat_STRING10;
    USER     : oscat_STRING32;
    PASSWORD : oscat_STRING32;
    DOMAIN   : oscat_STRING80;
    PORT     : WORD;
    PATH     : oscat_STRING80;
    QUERY    : oscat_STRING250;
    ANCHOR   : oscat_STRING40;
    HEADER   : oscat_STRING160;
    END_STRUCT;
END_TYPE

FUNCTION_BLOCK STRING_TO_URL_Block

	VAR_INPUT
		STR :	oscat_STRING250;
		DEFAULT_PROTOCOL :	oscat_STRING20 := 'http';
		DEFAULT_PATH :	oscat_STRING80 := '/';
	END_VAR

	VAR_OUTPUT
		STRING_TO_URL :	oscat_url;
	END_VAR

	VAR
		pos :	INT;
		pos2 :	INT;
		temp :	STRING;
		x :	oscat_STRING250;
	END_VAR

	IF EQ_STRING(STR,'') THEN
		RETURN;
	END_IF;

	pos := FIND(STR, '://');
	IF pos > 0 THEN
		STRING_TO_URL.PROTOCOL := LEFT(STR, pos - 1);
		x := RIGHT(STR, LEN(STR) - pos - 2);
	ELSE
		x := STR;
		STRING_TO_URL.PROTOCOL := DEFAULT_PROTOCOL;
	END_IF;

	pos := FIND(x, '@');
	IF pos > 0 THEN
		pos2 := FIND(x,':')+1;
		IF pos2 > 1 AND pos2 <= pos THEN
			STRING_TO_URL.USER := LEFT(x,pos2 - 2);
			STRING_TO_URL.PASSWORD := MID(x, pos - pos2, pos2);
		ELSE
			STRING_TO_URL.USER := LEFT(x, pos - 2);
			STRING_TO_URL.PASSWORD := '';
		END_IF;
		x := RIGHT(x, LEN(x) - pos);
	ELSE
		STRING_TO_URL.USER := '';
		STRING_TO_URL.PASSWORD := '';
	END_IF;

	pos := FIND(x, '#');
	IF pos > 0 THEN
		STRING_TO_URL.ANCHOR := RIGHT(x, LEN(x) - pos);
		x := LEFT(x, pos - 1);
	ELSE
		STRING_TO_URL.ANCHOR := '';
	END_IF;

	pos := FIND(x, '?');
	IF pos > 0 THEN
		STRING_TO_URL.QUERY := RIGHT(x, LEN(x) - pos);
		x := LEFT(x, pos - 1);
	ELSE
		STRING_TO_URL.QUERY := '';
	END_IF;

	pos := FIND(x, '/');
	IF pos > 0 THEN
		STRING_TO_URL.PATH := RIGHT(x, LEN(x) - pos + 1);
		x := LEFT(x, pos - 1);
	ELSE
		STRING_TO_URL.PATH := DEFAULT_PATH;
	END_IF;

	pos := FIND(x, ':');
	IF pos > 0 THEN
		temp := RIGHT(x, LEN(x) - pos);
		STRING_TO_URL.PORT := STRING_TO_WORD(temp);
		STRING_TO_URL.DOMAIN := LEFT(x, pos - 1);
	ELSE
		STRING_TO_URL.PORT := WORD#0;
		STRING_TO_URL.DOMAIN := x;
	END_IF;

END_FUNCTION_BLOCK

PROGRAM program0
	VAR
		STR :	oscat_STRING250;
		DEFAULT_PROTOCOL :	oscat_STRING20 := 'http';
		DEFAULT_PATH :	oscat_STRING80 := '/';
		STRING_TO_URL :	oscat_url;

		func_block : STRING_TO_URL_Block;
	END_VAR
	func_block.STR := STR;
	func_block.DEFAULT_PROTOCOL := DEFAULT_PROTOCOL;
	func_block.DEFAULT_PATH := DEFAULT_PATH;

	func_block();
  	STRING_TO_URL  := func_block.STRING_TO_URL;
END_PROGRAM

CONFIGURATION Config0
	RESOURCE Res0 ON PLC
		TASK task0(INTERVAL := T#20ms,PRIORITY := 0);
		PROGRAM instance0 WITH task0 : program0;
	END_RESOURCE
END_CONFIGURATION

(* ---- SUN_POS.ST ---- *)
FUNCTION FLOOR2 : DINT
	VAR_INPUT
		x : REAL;
	END_VAR

	FLOOR2 := REAL_TO_DINT(X);
	IF DINT_TO_REAL(FLOOR2) > X THEN
		FLOOR2 := FLOOR2 - DINT#1;
	END_IF;

END_FUNCTION

FUNCTION MODR:REAL

	VAR_INPUT
		IN :	REAL;
		DIVI :	REAL;
	END_VAR

	IF divi = 0.0 THEN
		MODR := 0.0;
	ELSE
		MODR := in - DINT_TO_REAL(FLOOR2(in / divi)) * divi;
	END_IF;

END_FUNCTION

FUNCTION RAD:REAL

	VAR_INPUT
		DEGG :	REAL;
	END_VAR

	RAD := MODR(0.0174532925199433 * DEGG , 6.283185307179586476);

END_FUNCTION

FUNCTION REFRACTION:REAL

	VAR_INPUT
		ELEV :	REAL;
	END_VAR

	VAR
		tmp :	REAL;
	END_VAR

	tmp := LIMIT(-1.9, elev, 80.0);
	REFRACTION := 0.0174532925199433 / TAN(0.0174532925199433 * (tmp + 10.3 / (tmp + 5.11)));

END_FUNCTION

FUNCTION TOD_TO_REAL2:REAL
	VAR_INPUT
		IN :	UDINT;
	END_VAR
	TOD_TO_REAL2 := UDINT_TO_REAL(IN);
END_FUNCTION

FUNCTION DEG:REAL

	VAR_INPUT
		X :	REAL;
	END_VAR

	DEG := MODR(57.29577951308232 * X, 360.0);
END_FUNCTION

FUNCTION DT_TO_TOD2:UDINT
	VAR_INPUT
		IN :	UDINT;
	END_VAR

	DT_TO_TOD2 := (IN MOD UDINT#86400) * UDINT#1000;
END_FUNCTION

FUNCTION_BLOCK SUN_POS

	VAR_INPUT
		LATITUDE :	REAL;
		LONGITUDE :	REAL;
		UTC :	UDINT;
	END_VAR

	VAR_OUTPUT
		B :	REAL;
		HR :	REAL;
	END_VAR

	VAR
		g :	REAL;
		a :	REAL;
		d :	REAL;
		h :	REAL;
		t1 :	REAL;
		n :	REAL;
		e :	REAL;
		c :	REAL;
		tau :	REAL;
		sin_d :	REAL;
		rlat :	REAL;
		sin_lat :	REAL;
		cos_lat :	REAL;
		cos_tau :	REAL;
		cos_d :	REAL;
		MATH_PI :	REAL := 3.14159265358979323846264338327950288;
		MATH_PI2 :	REAL := 6.28318530717958647692528676655900576;
	END_VAR

	n := UDINT_TO_REAL(UTC - UDINT#946728000) * 0.000011574074074074;
	g :=MODR(6.240040768 + 0.01720197 * n, MATH_PI2);
	d := MODR(4.89495042 + 0.017202792 * n, MATH_PI2) + 0.033423055 * SIN(g) + 0.000349066 * SIN(2.0*g);
	e := 0.409087723 - 0.000000006981317008 * n;
	cos_d := COS(d);
	sin_d := SIN(d);
	a := ATAN(COS(e) * sin_d / cos_d);
	IF cos_d < 0.0 THEN a := a + MATH_PI; END_IF;
	c := ASIN(SIN(e) * sin_d);

	(* also here we must be very careful utc is from 1.1.1970 for step7 the formula must change *)
	tau := RAD(MODR(6.697376 + (n - 0.25) * 0.0657098245037645 + TOD_TO_REAL2(DT_TO_TOD2(utc)) * 0.0000002785383333, 24.0) * 15.0 + longitude) - a;
	rlat := RAD(latitude);
	sin_lat := SIN(rlat);
	cos_lat := COS(rlat);
	cos_tau := COS(tau);
	t1 := cos_tau * sin_lat - TAN(c) * cos_lat;
	B := ATAN(SIN(tau) / t1);
	IF t1 < 0.0 THEN B := B + MATH_PI2; ELSE B := B + MATH_PI; END_IF;
	B := DEG(MODR(B, MATH_PI2));
	h := DEG(ASIN(COS(C) * cos_tau * cos_lat +SIN(c) * sin_lat));
	IF h > 180.0 THEN h := h - 360.0; END_IF;
	(* consider refraction *)
	HR := h + REFRACTION(h);
END_FUNCTION_BLOCK

PROGRAM program0
  VAR
	LATITUDE :	REAL;
	LONGITUDE :	REAL;
	UTC :	UDINT;
	B :	REAL;
	HR :	REAL;
	func_block : SUN_POS;
  END_VAR
	func_block.LATITUDE  :=LATITUDE ;
	func_block.LONGITUDE  :=LONGITUDE ;
	func_block.UTC  :=UTC ;
	func_block();
	B := func_block.B;
	HR := func_block.HR;
END_PROGRAM

CONFIGURATION Config0
	RESOURCE Res0 ON PLC
		TASK task0(INTERVAL := T#20ms,PRIORITY := 0);
		PROGRAM instance0 WITH task0 : program0;
	END_RESOURCE
END_CONFIGURATION

(* ---- SUN_TIME.ST ---- *)
FUNCTION RAD:REAL
	VAR_INPUT
		X:	REAL;
	END_VAR

	RAD := MODR(0.0174532925199433 * X , 6.283185307179586476);
END_FUNCTION

FUNCTION _REAL_TO_UDINT:UDINT

	VAR_INPUT
		X :	REAL;
	END_VAR

	IF REAL_TO_UDINT(0.5) = UDINT#1 THEN
		_REAL_TO_UDINT := REAL_TO_UDINT(x);
	ELSIF X > 0.0 THEN
		_REAL_TO_UDINT := REAL_TO_UDINT(x+0.5);
	ELSIF X < 0.0 THEN
		_REAL_TO_UDINT := REAL_TO_UDINT(x-0.5);
	ELSE
		_REAL_TO_UDINT := UDINT#0;
  	END_IF;
END_FUNCTION

FUNCTION HOUR_TO_TIME:TIME

	VAR_INPUT
		IN :	REAL;
	END_VAR

	hour_to_time := UDINT_TO_TIME(_REAL_TO_UDINT(IN * 3600000.0));
END_FUNCTION

FUNCTION TIME_TO_UDINT2:UDINT
	VAR_INPUT
		X :	TIME;
	END_VAR

	TIME_TO_UDINT2 := DINT_TO_UDINT(TIME_TO_DINT(X));
END_FUNCTION

FUNCTION FLOOR2 : DINT
	VAR_INPUT
		x : REAL;
	END_VAR

	FLOOR2 := REAL_TO_DINT(X);
	IF DINT_TO_REAL(FLOOR2) > X THEN
		FLOOR2 := FLOOR2 - DINT#1;
	END_IF;
END_FUNCTION

FUNCTION MODR:REAL

	VAR_INPUT
		IN :	REAL;
		DIVI :	REAL;
	END_VAR

	IF divi = 0.0 THEN
		MODR := 0.0;
	ELSE
		MODR := in - DINT_TO_REAL(FLOOR2(in / divi)) * divi;
	END_IF;

END_FUNCTION

FUNCTION DEG:REAL

	VAR_INPUT
		X :	REAL;
	END_VAR

	DEG := MODR(57.29577951308232 * X, 360.0);
END_FUNCTION

FUNCTION HOUR_TO_TOD:UDINT
	VAR_INPUT
		IN :	REAL;
	END_VAR

	hour_to_tod := _REAL_TO_UDINT(IN * 3600000.00);
END_FUNCTION

FUNCTION DAY_OF_YEAR:INT
	VAR_INPUT
		IDATE :	DATE;
	END_VAR

	DAY_OF_YEAR := UDINT_TO_INT((DATE_TO_UDINT(idate) / UDINT#86400) MOD UDINT#1461);
	IF DAY_OF_YEAR > 729 THEN
		IF DAY_OF_YEAR > 1095 THEN DAY_OF_YEAR := DAY_OF_YEAR - 1095; ELSE DAY_OF_YEAR := DAY_OF_YEAR - 729; END_IF;
	ELSIF DAY_OF_YEAR > 364 THEN
		DAY_OF_YEAR := DAY_OF_YEAR - 364;
	ELSE
		DAY_OF_YEAR := DAY_OF_YEAR + 1;
	END_IF;
END_FUNCTION

FUNCTION SUN_MIDDAY:UDINT
	VAR_INPUT
		LON :	REAL;
		UTC :	DATE;
	END_VAR

	VAR
		T :	REAL;
		OFFSET :	REAL;
	END_VAR

	T := INT_TO_REAL(DAY_OF_YEAR(utc));
	OFFSET := -0.1752 * SIN(0.033430 * T + 0.5474) - 0.1340 * SIN(0.018234 * T - 0.1939);
	SUN_MIDDAY := HOUR_TO_TOD(12.0 - OFFSET - lon * 0.0666666666666);
END_FUNCTION

FUNCTION_BLOCK SUN_TIME_Block

	VAR_INPUT
		LATITUDE :	REAL;
		LONGITUDE :	REAL;
		UTC :	DATE;
		H :	REAL := -0.83333333333;
	END_VAR

	VAR_OUTPUT
		MIDDAY :	UDINT;
		SUN_RISE :	UDINT;
		SUN_SET :	UDINT;
		SUN_DECLINATION :	REAL;
	END_VAR

	VAR
		DK :	REAL;
		delta :	UDINT;
		B :	REAL;
	END_VAR

	B := latitude * 0.0174532925199433;
	MIDDAY := SUN_MIDDAY(longitude, utc);
	DK := 0.40954 * SIN(0.0172 * (INT_TO_REAL(DAY_OF_YEAR(utc)) - 79.35));
	sun_declination := DEG(DK);
	IF sun_declination > 180.0 THEN sun_declination := sun_declination - 360.0; END_IF;
	sun_declination := 90.0 - LATITUDE + sun_declination;
	delta := TIME_TO_UDINT2(HOUR_TO_TIME(ACOS((SIN(RAD(H)) - SIN(B) * SIN(DK)) / (COS(B) * COS(DK))) * 3.819718632));
	sun_rise := MIDDAY - delta;
	sun_set := MIDDAY + delta;
END_FUNCTION_BLOCK

PROGRAM program0
  VAR
	LATITUDE :	REAL;
	LONGITUDE :	REAL;
	UTC :	DATE;
	H :	REAL := -0.83333333333;
	MIDDAY :	UDINT;
	SUN_RISE :	UDINT;
	SUN_SET :	UDINT;
	SUN_DECLINATION :	REAL;
	func_block : SUN_TIME_Block;
  END_VAR
	func_block.LATITUDE := LATITUDE;
	func_block.LONGITUDE := LONGITUDE;
	func_block.UTC := UTC;
	func_block.H := H;
	func_block();
	MIDDAY := func_block.MIDDAY;
	SUN_RISE := func_block.SUN_RISE;
	SUN_SET := func_block.SUN_SET;
	SUN_DECLINATION := func_block.SUN_DECLINATION;

END_PROGRAM

CONFIGURATION Config0

	RESOURCE Res0 ON PLC
		TASK task0(INTERVAL := T#20ms,PRIORITY := 0);
		PROGRAM instance0 WITH task0 : program0;
	END_RESOURCE

END_CONFIGURATION

(* ---- SW_RECONFIG.ST ---- *)
FUNCTION_BLOCK SW_RECONFIG_Block

	VAR_INPUT
		IN :	BOOL;
		TD :	TIME;
		TR :	TIME;
	END_VAR

	VAR_OUTPUT
		Q :	BOOL;
	END_VAR

	VAR
		T1 :	TON;
		T2 :	TON;
		INV :	BOOL;
	END_VAR

	t1(in := IN, PT := TD);

	IF tr > t#0s THEN
		Q := t1.Q XOR inv;
		T2(in := Q, pt := TR);
		IF T2.Q THEN INV := NOT INV; END_IF;
	ELSE
		Q := t1.Q;
	END_IF;

END_FUNCTION_BLOCK

PROGRAM program0
	VAR
		IN :	BOOL;
		TD :	TIME;
		TR :	TIME;
		Q :	BOOL;

		func_block : SW_RECONFIG_Block;
	END_VAR
	func_block.IN := IN;
	func_block.TD := TD;
	func_block.TR := TR ;

	func_block();
	Q  := func_block.Q;

END_PROGRAM

CONFIGURATION Config0
	RESOURCE Res0 ON PLC
		TASK task0(INTERVAL := T#20ms,PRIORITY := 0);
		PROGRAM instance0 WITH task0 : program0;
	END_RESOURCE
END_CONFIGURATION

(* ---- SWITCH_I.ST ---- *)
FUNCTION UDINT_TO_TIME2:TIME

	VAR_INPUT
		IN :	UDINT;
	END_VAR

	UDINT_TO_TIME2 := DINT_TO_TIME(UDINT_TO_DINT(IN));

END_FUNCTION

FUNCTION_BLOCK T_PLC_MS_block
	VAR_OUTPUT
		T_PLC_MS :	UDINT;
	END_VAR

	VAR_EXTERNAL
		PLC_TICKS_PER_SEC :	INT;
		PLC_SYS_TICK_CNT :	DINT;
	END_VAR

	VAR
		debug :	BOOL;(*Debug-Mode ON / OFF*)
		N :	INT;(*Debug-Faktor*)
		Offset :	UDINT;(*Debug-Offset*)
		temp :	DWORD := DWORD#1;(*Debug-Offset*)
		mode :	BOOL;(*modus*)
		faktor :	UDINT;(*Systemtakt-Faktor*)
		init :	BOOL;
		v_plc_ticks_per_sec :	UDINT;
		base :	UDINT := UDINT#1000;
	END_VAR

	IF init = FALSE THEN
		v_plc_ticks_per_sec := INT_TO_UDINT(PLC_TICKS_PER_SEC);
		IF v_plc_ticks_per_sec = UDINT#1024 THEN
			faktor := UDINT#1;
			mode := FALSE;
		ELSIF v_plc_ticks_per_sec > UDINT#0 THEN
			IF v_plc_ticks_per_sec <= base THEN
				faktor := base / v_plc_ticks_per_sec;
				mode := FALSE;
			ELSE
				faktor := v_plc_ticks_per_sec / base;
				mode := TRUE;
			END_IF;
		ELSE
			faktor := UDINT#1;
		END_IF;
		init := TRUE;
	END_IF;

	IF mode THEN
		T_PLC_MS := DINT_TO_UDINT(PLC_SYS_TICK_CNT) / faktor;
	ELSE
		T_PLC_MS := DINT_TO_UDINT(PLC_SYS_TICK_CNT) * faktor;
	END_IF;

	IF debug THEN
		T_PLC_MS := (DWORD_TO_UDINT(SHL(UDINT_TO_DWORD(T_PLC_MS),N) OR SHL(temp,N)) - UDINT#1) + Offset;
	END_IF;

END_FUNCTION_BLOCK

FUNCTION_BLOCK SWITCH_I_Block

	VAR_INPUT
		SET :	BOOL;
		IN :	BOOL;
		RST :	BOOL;
		T_DEBOUNCE :	TIME := T#10ms;
		T_RECONFIG :	TIME := T#1s;
		T_ON_MAX :	TIME := T#0h;
	END_VAR

	VAR_OUTPUT
		Q :	BOOL := FALSE;
	END_VAR

	VAR
		state :	BYTE := BYTE#0;
		edge :	BOOL := FALSE;
		_r_edge :	BOOL := FALSE;
		T_on :	TIME;
		tx :	TIME;
		T_PLC_MS :	T_PLC_MS_Block;
	END_VAR

	T_PLC_MS();
	tx:= UDINT_TO_TIME(T_PLC_MS.T_PLC_MS);

	IF set AND NOT rst THEN
		Q := TRUE;
		T_on := tx;
	ELSIF rst THEN
		Q := FALSE;
	ELSIF (in XOR edge) AND NOT (state = BYTE#1) THEN
		state := BYTE#1;
		T_on := Tx;
	ELSIF (state = BYTE#1) AND (Tx - t_debounce >= T_on) THEN
		state := BYTE#2;
		IF _r_edge XOR in THEN Q := NOT Q;
	END_IF;
	ELSIF state = BYTE#2 AND Tx - t_reconfig >= T_on THEN
		_r_edge := in;
	END_IF;
	IF Q AND T_on_max > t#0ms AND Tx >= T_on + T_on_max THEN
		Q := FALSE;
	END_IF;
	edge := in;

END_FUNCTION_BLOCK

PROGRAM program0
	VAR
		SET :	BOOL;
		IN :	BOOL;
		RST :	BOOL;
		T_DEBOUNCE :	TIME := T#10ms;
		T_RECONFIG :	TIME := T#1s;
		T_ON_MAX :	TIME := T#0h;
		Q :	BOOL := FALSE;

		func_block : SWITCH_I_Block;
	END_VAR
	func_block.SET := SET;
	func_block.IN := IN;
	func_block.RST := RST ;
	func_block.T_DEBOUNCE := T_DEBOUNCE ;
	func_block.T_RECONFIG := T_RECONFIG ;
	func_block.T_ON_MAX := T_ON_MAX ;

	func_block();
	Q  := func_block.Q;
END_PROGRAM

CONFIGURATION Config0
	VAR_GLOBAL
		PLC_TICKS_PER_SEC :	INT;
		PLC_SYS_TICK_CNT :	DINT;
	END_VAR
  	RESOURCE Res0 ON PLC
    	TASK task0(INTERVAL := T#20ms,PRIORITY := 0);
    	PROGRAM instance0 WITH task0 : program0;
  	END_RESOURCE
END_CONFIGURATION

(* ---- SWITCH_X.ST ---- *)
FUNCTION_BLOCK SWITCH_X_Block

	VAR_INPUT
		IN1 :	BOOL;
		IN2 :	BOOL;
		IN3 :	BOOL;
		IN4 :	BOOL;
		IN5 :	BOOL;
		IN6 :	BOOL;
		T_DEBOUNCE :	TIME := T#50ms;
	END_VAR

	VAR_OUTPUT
		Q1 :	BOOL;
		Q2 :	BOOL;
		Q3 :	BOOL;
		Q4 :	BOOL;
		Q5 :	BOOL;
		Q6 :	BOOL;
		Q31 :	BOOL;
		Q41 :	BOOL;
		Q51 :	BOOL;
		Q61 :	BOOL;
		Q32 :	BOOL;
		Q42 :	BOOL;
		Q52 :	BOOL;
		Q62 :	BOOL;
	END_VAR

	VAR
		INIT :	BOOL;
		T1 :	TOF;
		T2 :	TOF;
		T3 :	TOF;
		T4 :	TOF;
		T5 :	TOF;
		T6 :	TOF;
		tx :	TIME;
		x1 :	BOOL;
		x2 :	BOOL;
		E1 :	BOOL;
		E2 :	BOOL;
	END_VAR

	IF NOT init THEN
		init := TRUE;
		IF t_debounce < t#50ms THEN tx := t#50ms; ELSE tx := t_debounce; END_IF;
		T1(PT := Tx);
		T2(PT := Tx);
		T3(PT := Tx);
		T4(PT := Tx);
		T5(PT := Tx);
		T6(PT := Tx);
	ELSE
		Q1 := FALSE;
		Q2 := FALSE;
		Q3 := FALSE;
		Q4 := FALSE;
		Q5 := FALSE;
		Q6 := FALSE;
		Q31 := FALSE;
		Q41 := FALSE;
		Q51 := FALSE;
		Q61 := FALSE;
		Q32 := FALSE;
		Q42 := FALSE;
		Q52 := FALSE;
		Q62 := FALSE;
	END_IF;

		T1(IN := IN1);
		T2(IN := IN2);
		T3(IN := IN3);
		T4(IN := IN4);
		T5(IN := IN5);
		T6(IN := IN6);

	IF t1.Q AND NOT E1 THEN X1 := TRUE; END_IF;
	IF t2.Q AND NOT E2 THEN X2 := TRUE; END_IF;

	IF t1.Q THEN
		IF t3.q THEN
			q31 := TRUE;
			X1 := FALSE;
		ELSIF t4.q THEN
			q41 := TRUE;
			X1 := FALSE;
		ELSIF t5.q THEN
			q51 := TRUE;
			X1 := FALSE;
		ELSIF t6.q THEN
			q61 := TRUE;
			X1 := FALSE;
		END_IF;
	ELSIF t2.Q THEN
		IF t3.q THEN
			q32 := TRUE;
			X2 := FALSE;
		ELSIF t4.q THEN
			q42 := TRUE;
			X2 := FALSE;
		ELSIF t5.q THEN
			q52 := TRUE;
			X2 := FALSE;
		ELSIF t6.q THEN
			q62 := TRUE;
			X2 := FALSE;
		END_IF;
	ELSIF NOT T1.Q AND E1 AND X1 THEN
		Q1 := TRUE;
		X1 := FALSE;
	ELSIF NOT T2.Q AND E2 AND X2 THEN
		Q2 := TRUE;
		X2 := FALSE;
	ELSIF T3.Q THEN
		Q3 := TRUE;
	ELSIF T4.Q THEN
		Q4 := TRUE;
	ELSIF T5.Q THEN
		Q5 := TRUE;
	ELSIF T6.Q THEN
		Q6 := TRUE;
	END_IF;

	E1 := T1.Q;
	E2 := T2.Q;
END_FUNCTION_BLOCK

PROGRAM program0
	VAR
		IN1 :	BOOL;
		IN2 :	BOOL;
		IN3 :	BOOL;
		IN4 :	BOOL;
		IN5 :	BOOL;
		IN6 :	BOOL;
		T_DEBOUNCE :	TIME := T#50ms;
		Q1 :	BOOL;
		Q2 :	BOOL;
		Q3 :	BOOL;
		Q4 :	BOOL;
		Q5 :	BOOL;
		Q6 :	BOOL;
		Q31 :	BOOL;
		Q41 :	BOOL;
		Q51 :	BOOL;
		Q61 :	BOOL;
		Q32 :	BOOL;
		Q42 :	BOOL;
		Q52 :	BOOL;
		Q62 :	BOOL;

		func_block : SWITCH_X_Block;
	END_VAR
	func_block.IN1 := IN1;
	func_block.IN2 := IN2;
	func_block.IN3 := IN3 ;
	func_block.IN4 := IN4;
	func_block.IN5 := IN5;
	func_block.IN6 := IN6 ;
	func_block.T_DEBOUNCE := T_DEBOUNCE;

	func_block();
	Q1  := func_block.Q1;
	Q2  := func_block.Q2;
	Q3  := func_block.Q3;
	Q4  := func_block.Q4;
	Q5  := func_block.Q5;
	Q6  := func_block.Q6;
	Q31  := func_block.Q31;
	Q41  := func_block.Q41;
	Q51  := func_block.Q51;
	Q61  := func_block.Q61;
	Q32  := func_block.Q32;
	Q42  := func_block.Q42;
	Q52  := func_block.Q52;
	Q62  := func_block.Q62;

END_PROGRAM

CONFIGURATION Config0
	RESOURCE Res0 ON PLC
		TASK task0(INTERVAL := T#20ms,PRIORITY := 0);
		PROGRAM instance0 WITH task0 : program0;
	END_RESOURCE
END_CONFIGURATION

(* ---- SYS_LOG.ST ---- *)
FUNCTION_BLOCK SYS_LOG

  VAR_EXTERNAL

  END_VAR

  VAR

  END_VAR

  VAR_IN_OUT
    IP_C :	oscat_IP_C;
    S_BUF :	oscat_NETWORK_BUFFER;
    R_BUF :	oscat_NETWORK_BUFFER;
  END_VAR

  VAR_INPUT
    ACTIVATE :	BOOL;
    LDT :	UDINT;
    SERVER_IP4 :	DWORD;
    PORT :	WORD;
    FACILITY :	BYTE;
    SEVERITY :	BYTE;
    TAG :	oscat_STRING32;
    HOSTNAME :	STRING;
    MESSAGE :	oscat_STRING250;
    OPTION :	BYTE;
  END_VAR

  VAR_OUTPUT
    DONE_P :	BOOL;
    ERROR :	DWORD;
  END_VAR

  VAR
    IP_FIFO :	IP_FIFO;
    _STRING_TO_BUFFER :	_STRING_TO_BUFFER_NW;
    DT_TO_STRF :	DT_TO_STRF;
    ip_state :	BYTE;
    ip_id :	BYTE;
    activate_last :	BOOL;
    state :	INT;
    s1 :	oscat_STRING20;
    i :	INT;
  END_VAR

  CASE state OF
  00:
    IF ACTIVATE AND NOT activate_last THEN
      state := 10;
      ERROR := DWORD#0;
      ip_state := BYTE#1;
    END_IF;
    DONE_P := FALSE;

  10:
    IF ip_state = BYTE#3 THEN
      i := 0;

      IF (OPTION AND BYTE#0000_0001) = BYTE#00 THEN
        s1:=REPLACE('<P>',BYTE_TO_STRING(SHL_BYTE(FACILITY,3) OR (SEVERITY AND BYTE#0000_0111),'%u'),1,2);
      ELSE
        s1 := '';
      END_IF;

      IF (OPTION AND BYTE#0000_0010) = BYTE#00 THEN
        DT_TO_STRF(DTI:=LDT,MS:=0,FMT:='#E #W #N:#R:#T ',LANG:=1);
        s1 := CONCAT(s1,DT_TO_STRF.DT_TO_STRF);

        _STRING_TO_BUFFER(str:=s1,pos:=i,size:=UINT#1024,pt:=S_BUF.BUFFER);
        S_BUF.BUFFER:=_STRING_TO_BUFFER.pt;

        i := i + LEN(s1);

        _STRING_TO_BUFFER(str:=HOSTNAME,pos:=i,size:=UINT#1024,pt:=S_BUF.BUFFER);
        S_BUF.BUFFER:=_STRING_TO_BUFFER.pt;

        i := i + LEN(HOSTNAME);
        S_BUF.BUFFER[i] := BYTE#32;
        i := i + 1;

        _STRING_TO_BUFFER(str:=TAG,pos:=i,size:=UINT#1024,pt:=S_BUF.BUFFER);
        S_BUF.BUFFER:=_STRING_TO_BUFFER.pt;

        i := i + LEN(TAG);
        S_BUF.BUFFER[i] := BYTE#32;
        i := i + 1;
      END_IF;

      _STRING_TO_BUFFER(str:=MESSAGE,pos:=i,size:=UINT#1024,pt:=S_BUF.BUFFER);
      S_BUF.BUFFER:=_STRING_TO_BUFFER.pt;

      i := i + LEN(MESSAGE);

      IF (OPTION AND BYTE#0000_0100) > BYTE#00 THEN
        S_BUF.BUFFER[i] := BYTE#13;
        i := i + 1;
        S_BUF.BUFFER[i] := BYTE#10;
        i := i + 1;
      END_IF;

      state := 30;

      IF (OPTION AND BYTE#2#0000_1000) > BYTE#00 THEN
        IP_C.C_MODE := BYTE#0;
      ELSE
        IP_C.C_MODE := BYTE#1;
      END_IF;

      IF PORT = WORD#0 THEN
        IF IP_C.C_MODE = BYTE#0 THEN
          IP_C.C_PORT := WORD#1468;
      ELSE
          IP_C.C_PORT := WORD#514;
        END_IF;
      ELSE
        IP_C.C_PORT := PORT;
    END_IF;

      IP_C.C_IP       := SERVER_IP4;
      IP_C.C_ENABLE   := TRUE;
      IP_C.TIME_RESET := TRUE;
      IP_C.R_OBSERVE  := FALSE;
      S_BUF.SIZE      := INT_TO_UINT(i);
      R_BUF.SIZE      := UINT#0;
    END_IF;

  30:
    IF IP_C.ERROR <> DWORD#00 THEN
      ERROR := IP_C.ERROR;
      state := 0;

    ELSIF S_BUF.SIZE = UINT#0 THEN
      DONE_P := TRUE;
      state := 0;
    END_IF;

    IF state = 0 THEN
      ip_state := BYTE#4;
    END_IF;

  END_CASE;

  activate_last := ACTIVATE;

  IP_FIFO(FIFO:=IP_C.FIFO,state:=IP_STATE,ID:=ip_id);
  IP_C.FIFO := IP_FIFO.FIFO;
  ip_state := IP_FIFO.STATE;
  ip_id := IP_FIFO.ID;

END_FUNCTION_BLOCK

(* ---- T_AVG24.ST ---- *)
TYPE
  oscat_T_AVG24         	  : ARRAY [0..47]   OF INT;
END_TYPE

FUNCTION_BLOCK T_PLC_MS_block
	VAR_OUTPUT
		T_PLC_MS :	UDINT;
	END_VAR

	VAR_EXTERNAL
		PLC_TICKS_PER_SEC :	INT;
		PLC_SYS_TICK_CNT :	DINT;
	END_VAR

	VAR
		debug :	BOOL;(*Debug-Mode ON / OFF*)
		N :	INT;(*Debug-Faktor*)
		Offset :	UDINT;(*Debug-Offset*)
		temp :	DWORD := DWORD#1;(*Debug-Offset*)
		mode :	BOOL;(*modus*)
		faktor :	UDINT;(*Systemtakt-Faktor*)
		init :	BOOL;
		v_plc_ticks_per_sec :	UDINT;
		base :	UDINT := UDINT#1000;
	END_VAR

	IF init = FALSE THEN
		v_plc_ticks_per_sec := INT_TO_UDINT(PLC_TICKS_PER_SEC);
		IF v_plc_ticks_per_sec = UDINT#1024 THEN
			faktor := UDINT#1;
			mode := FALSE;
		ELSIF v_plc_ticks_per_sec > UDINT#0 THEN
			IF v_plc_ticks_per_sec <= base THEN
				faktor := base / v_plc_ticks_per_sec;
				mode := FALSE;
			ELSE
				faktor := v_plc_ticks_per_sec / base;
				mode := TRUE;
			END_IF;
		ELSE
			faktor := UDINT#1;
		END_IF;
		init := TRUE;
	END_IF;

	IF mode THEN
		T_PLC_MS := DINT_TO_UDINT(PLC_SYS_TICK_CNT) / faktor;
	ELSE
		T_PLC_MS := DINT_TO_UDINT(PLC_SYS_TICK_CNT) * faktor;
	END_IF;

	IF debug THEN
		T_PLC_MS := (DWORD_TO_UDINT(SHL(UDINT_TO_DWORD(T_PLC_MS),N) OR SHL(temp,N)) - UDINT#1) + Offset;
	END_IF;

END_FUNCTION_BLOCK

FUNCTION_BLOCK FILTER_I_Block
	VAR_INPUT
		X :	INT;
		T :	TIME;
	END_VAR

	VAR_OUTPUT
		Y :	INT;
	END_VAR

	VAR
		Yi :	DINT;
		last :	UDINT;
		tx :	UDINT;
		init :	BOOL;
		T_PLC_MS :	T_PLC_MS_block;
	END_VAR

	T_PLC_MS();
	tx:= T_PLC_MS.T_PLC_MS;

	IF NOT init OR T = t#0s THEN
		init := TRUE;
		Yi := INT_TO_DINT(X) * DINT#1000;
	ELSE
		Yi := Yi + INT_TO_DINT(X - Y) * UDINT_TO_DINT(tx - last) * DINT#1000 / TIME_TO_DINT(T);
	END_IF;
	last := tx;
	Y := DINT_TO_INT(yi / DINT#1000);

END_FUNCTION_BLOCK

FUNCTION TIME_TO_UDINT2:UDINT
	VAR_INPUT
		X :	TIME;
	END_VAR

	TIME_TO_UDINT2 := DINT_TO_UDINT(TIME_TO_DINT(X));
END_FUNCTION

FUNCTION INC1:INT

	VAR_INPUT
		X :	INT;
		N :	INT;
	END_VAR

	IF X >= N - 1 THEN
		INC1 := 0;
	ELSE
		INC1 := X + 1;
	END_IF;
END_FUNCTION

FUNCTION_BLOCK T_AVG24_Block

	VAR_INPUT
		TS :	INT;
		DTI :	UDINT;
		RST :	BOOL;
		T_FILTER :	TIME := T#10m;
		SCALE :	REAL := 1.0;
		OFS :	REAL;
	END_VAR

	VAR_OUTPUT
		TA :	REAL;
		_TP :	BOOL;
	END_VAR

	VAR_IN_OUT
		T24 :	REAL;
		T24_MAX :	REAL;
		T24_MIN :	REAL;
	END_VAR

	VAR
		samples :	oscat_T_AVG24;
		pos :	INT;
		init :	BOOL;
		sum :	DINT;
		last :	UDINT;
		tmp_maxxx :	INT;
		tmp_min :	INT;
		i :	INT;
		ft1 :	FILTER_I_Block;
	END_VAR

	ft1(X := TS, T := T_FILTER);

	IF rst OR NOT init THEN
		init := TRUE;
		IF T24 = -1000.0 THEN t24 := INT_TO_REAL(ft1.Y) * 0.1; END_IF;
		FOR pos := 0 TO 47 DO
			samples[pos] := REAL_TO_INT(T24 * 10.0);
		END_FOR;
		pos := 0;
		sum := INT_TO_DINT(samples[0]) * DINT#48;
		TA := (INT_TO_REAL(ft1.Y) * 0.1 + OFS) * SCALE;
		T24 := (DINT_TO_REAL(sum) * 0.00208333333333 + OFS) * SCALE;
		_TP := TRUE;
	ELSIF (dti / UDINT#60 MOD UDINT#30) = UDINT#0 AND DTI > last THEN
		last := DTI + TIME_TO_UDINT2(T#1m);
		sum := sum - INT_TO_DINT(samples[pos]);
		samples[pos] := ft1.Y;
		sum := sum + INT_TO_DINT(samples[pos]);
		pos := INC1(pos, 48);
		TA := (INT_TO_REAL(ft1.Y) * 0.1 + OFS) * SCALE;
		T24 := (DINT_TO_REAL(sum) * 0.00208333333333 + OFS) * SCALE;
		tmp_maxxx := -32000;
		tmp_min := 32000;
		FOR i := 0 TO 47 DO
			tmp_maxxx := MAX(tmp_maxxx, samples[i]);
			tmp_min := MIN(tmp_min, samples[i]);
		END_FOR;
		T24_MAX := (INT_TO_REAL(tmp_maxxx) * 0.1 + OFS) * SCALE;
		T24_MIN := (INT_TO_REAL(tmp_min) * 0.1 + OFS) * SCALE;
		_TP := TRUE;
	ELSE
		_TP := FALSE;
	END_IF;

END_FUNCTION_BLOCK

PROGRAM program0
	VAR
		TS :	INT;
		DTI :	UDINT;
		RST :	BOOL;
		T_FILTER :	TIME := T#10m;
		SCALE :	REAL := 1.0;
		OFS :	REAL;
		TA :	REAL;
		_TP :	BOOL;

		func_block : T_AVG24_Block;
	END_VAR
	func_block.TS := TS;
	func_block.DTI := DTI;
	func_block.RST := RST ;
	func_block.T_FILTER := T_FILTER;
	func_block.SCALE := SCALE;
	func_block.OFS := OFS ;

	func_block();
	TA  := func_block.TA;
	_TP  := func_block._TP;

END_PROGRAM

CONFIGURATION Config0
	VAR_GLOBAL
		PLC_TICKS_PER_SEC :	INT;
		PLC_SYS_TICK_CNT :	DINT;
	END_VAR
  	RESOURCE Res0 ON PLC
    	TASK task0(INTERVAL := T#20ms,PRIORITY := 0);
    	PROGRAM instance0 WITH task0 : program0;
  	END_RESOURCE
END_CONFIGURATION

(* ---- T_PLC_MS.ST ---- *)
FUNCTION_BLOCK T_PLC_MS_block

	VAR_OUTPUT
		T_PLC_MS :	UDINT;
	END_VAR

	VAR_EXTERNAL
		PLC_TICKS_PER_SEC :	INT;
		PLC_SYS_TICK_CNT :	DINT;
	END_VAR

	VAR
		debug :	BOOL;(*Debug-Mode ON / OFF*)
		N :	INT;(*Debug-Faktor*)
		Offset :	UDINT;(*Debug-Offset*)
		temp :	DWORD := DWORD#1;(*Debug-Offset*)
		mode :	BOOL;(*modus*)
		faktor :	UDINT;(*Systemtakt-Faktor*)
		init :	BOOL;
		v_plc_ticks_per_sec :	UDINT;
		base :	UDINT := UDINT#1000;
	END_VAR

	IF init = FALSE THEN
		v_plc_ticks_per_sec := INT_TO_UDINT(PLC_TICKS_PER_SEC);
		IF v_plc_ticks_per_sec = UDINT#1024 THEN
			faktor := UDINT#1;
			mode := FALSE;
		ELSIF v_plc_ticks_per_sec > UDINT#0 THEN
			IF v_plc_ticks_per_sec <= base THEN
				faktor := base / v_plc_ticks_per_sec;
				mode := FALSE;
			ELSE
				faktor := v_plc_ticks_per_sec / base;
				mode := TRUE;
			END_IF;
		ELSE
			faktor := UDINT#1;
		END_IF;
		init := TRUE;
	END_IF;

	IF mode THEN
		T_PLC_MS := DINT_TO_UDINT(PLC_SYS_TICK_CNT) / faktor;
	ELSE
		T_PLC_MS := DINT_TO_UDINT(PLC_SYS_TICK_CNT) * faktor;
	END_IF;

	IF debug THEN
		T_PLC_MS := (DWORD_TO_UDINT(SHL(UDINT_TO_DWORD(T_PLC_MS),N) OR SHL(temp,N)) - UDINT#1) + Offset;
	END_IF;

END_FUNCTION_BLOCK

PROGRAM program0

	VAR
		LocalOUT  : UDINT;
		func_block : T_PLC_MS_block;
  	END_VAR

	func_block();
	LocalOUT := func_block.T_PLC_MS;

END_PROGRAM

CONFIGURATION Config0

	VAR_GLOBAL
		PLC_TICKS_PER_SEC :	INT;
		PLC_SYS_TICK_CNT :	DINT;
	END_VAR

  	RESOURCE Res0 ON PLC
    	TASK task0(INTERVAL := T#20ms,PRIORITY := 0);
    	PROGRAM instance0 WITH task0 : program0;
  	END_RESOURCE

END_CONFIGURATION

(* ---- T_PLC_US.ST ---- *)
FUNCTION_BLOCK T_PLC_US_Block

	VAR_OUTPUT
		T_PLC_US :	UDINT;
	END_VAR

	VAR_EXTERNAL
		PLC_TICKS_PER_SEC :	INT;
		PLC_SYS_TICK_CNT :	DINT;
	END_VAR

	VAR
		debug :	BOOL;
		N :	INT;
		Offset :	UDINT;
		temp :	DWORD := DWORD#1;
		mode :	BOOL;
		faktor :	UDINT;
		init :	BOOL;
		v_plc_ticks_per_sec :	UDINT;
		base :	UDINT := UDINT#1000000;
	END_VAR

	IF init = FALSE THEN
		v_plc_ticks_per_sec := INT_TO_UDINT(PLC_TICKS_PER_SEC);
		IF v_plc_ticks_per_sec = UDINT#1024 THEN
			faktor := UDINT#1000;
			mode := FALSE;
		ELSIF v_plc_ticks_per_sec > UDINT#0 THEN
			IF v_plc_ticks_per_sec <= base THEN
				faktor := base / v_plc_ticks_per_sec;
				mode := FALSE;
			ELSE
				faktor := v_plc_ticks_per_sec / base;
				mode := TRUE;
			END_IF;
		ELSE
			faktor := UDINT#1;
		END_IF;
		init := TRUE;
	END_IF;

	IF mode THEN
		T_PLC_US := DINT_TO_UDINT(PLC_SYS_TICK_CNT) / faktor;
	ELSE
		T_PLC_US := DINT_TO_UDINT(PLC_SYS_TICK_CNT) * faktor;
	END_IF;

	IF debug THEN
		T_PLC_US := (DWORD_TO_UDINT(SHL(UDINT_TO_DWORD(T_PLC_US),N) OR SHL(temp,N)) - UDINT#1) + Offset;
	END_IF;

END_FUNCTION_BLOCK

PROGRAM program0

	VAR
		T_PLC_US  : UDINT;
		func_block : T_PLC_US_Block;
	END_VAR
		func_block();
		T_PLC_US := func_block.T_PLC_US;

END_PROGRAM

CONFIGURATION Config0

	VAR_GLOBAL
		PLC_TICKS_PER_SEC :	INT;
		PLC_SYS_TICK_CNT :	DINT;
	END_VAR

	RESOURCE Res0 ON PLC
		TASK task0(INTERVAL := T#20ms,PRIORITY := 0);
		PROGRAM instance0 WITH task0 : program0;
	END_RESOURCE

END_CONFIGURATION

(* ---- TANK_LEVEL.ST ---- *)
FUNCTION_BLOCK TONOF

	VAR_INPUT
		IN :	BOOL;
		T_ON :	TIME;
		T_OFF :	TIME;
	END_VAR

	VAR_OUTPUT
		Q :	BOOL;
	END_VAR

	VAR
		X :	TON;
		old :	BOOL;
		mode :	BOOL;
	END_VAR

	IF IN XOR old THEN
	X(IN := FALSE, PT := SEL_TIME(IN,T_OFF,T_ON));
	mode := IN;
	old := IN;
	END_IF;
	X(IN := TRUE);
	IF X.Q THEN Q := mode;END_IF;

END_FUNCTION_BLOCK

FUNCTION UDINT_TO_TIME2:TIME

	VAR_INPUT
		IN :	UDINT;
	END_VAR

	UDINT_TO_TIME2 := DINT_TO_TIME(UDINT_TO_DINT(IN));

END_FUNCTION

FUNCTION_BLOCK T_PLC_MS_block
	VAR_OUTPUT
		T_PLC_MS :	UDINT;
	END_VAR

	VAR_EXTERNAL
		PLC_TICKS_PER_SEC :	INT;
		PLC_SYS_TICK_CNT :	DINT;
	END_VAR

	VAR
		debug :	BOOL;(*Debug-Mode ON / OFF*)
		N :	INT;(*Debug-Faktor*)
		Offset :	UDINT;(*Debug-Offset*)
		temp :	DWORD := DWORD#1;(*Debug-Offset*)
		mode :	BOOL;(*modus*)
		faktor :	UDINT;(*Systemtakt-Faktor*)
		init :	BOOL;
		v_plc_ticks_per_sec :	UDINT;
		base :	UDINT := UDINT#1000;
	END_VAR

	IF init = FALSE THEN
		v_plc_ticks_per_sec := INT_TO_UDINT(PLC_TICKS_PER_SEC);
		IF v_plc_ticks_per_sec = UDINT#1024 THEN
			faktor := UDINT#1;
			mode := FALSE;
		ELSIF v_plc_ticks_per_sec > UDINT#0 THEN
			IF v_plc_ticks_per_sec <= base THEN
				faktor := base / v_plc_ticks_per_sec;
				mode := FALSE;
			ELSE
				faktor := v_plc_ticks_per_sec / base;
				mode := TRUE;
			END_IF;
		ELSE
			faktor := UDINT#1;
		END_IF;
		init := TRUE;
	END_IF;

	IF mode THEN
		T_PLC_MS := DINT_TO_UDINT(PLC_SYS_TICK_CNT) / faktor;
	ELSE
		T_PLC_MS := DINT_TO_UDINT(PLC_SYS_TICK_CNT) * faktor;
	END_IF;

	IF debug THEN
		T_PLC_MS := (DWORD_TO_UDINT(SHL(UDINT_TO_DWORD(T_PLC_MS),N) OR SHL(temp,N)) - UDINT#1) + Offset;
	END_IF;
END_FUNCTION_BLOCK

FUNCTION TIME_TO_UDINT2:UDINT
	VAR_INPUT
		X :	TIME;
	END_VAR

	TIME_TO_UDINT2 := DINT_TO_UDINT(TIME_TO_DINT(X));
END_FUNCTION

FUNCTION_BLOCK ACTUATOR_COIL_Block

	VAR_INPUT
		IN :	BOOL;
		SELF_ACT_CYCLE :	TIME := T#10d;
		SELF_ACT_TIME :	TIME := T#1s;
	END_VAR

	VAR_OUTPUT
		OUT :	BOOL;
		STATUS :	BYTE;
	END_VAR

	VAR
		last :	UDINT;
		init :	BOOL;
		tx :	UDINT;
		now :	UDINT;
		T_PLC_MS :	T_PLC_MS_Block;
	END_VAR

	T_PLC_MS();
	now := T_PLC_MS.T_PLC_MS;

	IF NOT init THEN
		last := now;
		init := TRUE;
	ELSIF IN THEN
		OUT := TRUE;
		STATUS := BYTE#101;
		LAST := now;
	ELSE
		OUT := FALSE;
		STATUS := BYTE#100;
		tx := now - last;
		IF (self_act_cycle > T#0s) AND (tx >= TIME_TO_UDINT2(self_act_cycle)) THEN
			OUT := TRUE;
			STATUS := BYTE#102;
			IF tx >= TIME_TO_UDINT2(self_act_cycle + self_act_time) THEN
				last := now;
				OUT := FALSE;
				STATUS := BYTE#100;
			END_IF;
		END_IF;
	END_IF;

END_FUNCTION_BLOCK

FUNCTION_BLOCK TANK_LEVEL_Block

	VAR_INPUT
		LEVEL :	BOOL;
		LEAK :	BOOL;
		ACLR :	BOOL;
		MAX_VALVE_TIME :	TIME;
		LEVEL_DELAY_TIME :	TIME;
	END_VAR

	VAR_OUTPUT
		VALVE :	BOOL;
		ALARM :	BOOL;
		STATUS :	BYTE;
	END_VAR

	VAR
		cx :	ACTUATOR_COIL_Block;
		tn :	TON;
		tl :	TONOF;
		open :	BOOL;
	END_VAR

	tl(in := level, T_ON := level_delay_time, T_OFF := level_delay_time);
	open := tl.Q;

	IF ALARM THEN
		IF ACLR THEN
			ALARM := FALSE;
			STATUS := BYTE#101;
			cx(in := FALSE);
		END_IF;
		RETURN;
	ELSIF LEAK THEN
		cx(in := FALSE);
		ALARM := TRUE;
		STATUS := BYTE#1;
	ELSIF open THEN
		cx(in := TRUE);
		STATUS := BYTE#102;
	ELSE
		cx(in := FALSE);
		STATUS := BYTE#100;
	END_IF;

	tn(in := cx.out AND (MAX_VALVE_TIME > T#0s), PT := MAX_VALVE_TIME);
	IF tn.Q THEN
		ALARM := TRUE;
		STATUS := BYTE#2;
		cx(in := FALSE);
	END_IF;

	VALVE := cx.out;
END_FUNCTION_BLOCK

PROGRAM program0
	VAR
		LEVEL :	BOOL;
		LEAK :	BOOL;
		ACLR :	BOOL;
		MAX_VALVE_TIME :	TIME;
		LEVEL_DELAY_TIME :	TIME;
		VALVE :	BOOL;
		ALARM :	BOOL;
		STATUS :	BYTE;

		func_block : TANK_LEVEL_Block;
	END_VAR
	func_block.LEVEL := LEVEL;
	func_block.LEAK := LEAK;
	func_block.ACLR := ACLR ;
	func_block.MAX_VALVE_TIME := MAX_VALVE_TIME;
	func_block.LEVEL_DELAY_TIME := LEVEL_DELAY_TIME ;
	func_block();
	VALVE  := func_block.VALVE;
	ALARM  := func_block.ALARM;
	STATUS  := func_block.STATUS;
END_PROGRAM

CONFIGURATION Config0
	VAR_GLOBAL
		PLC_TICKS_PER_SEC :	INT;
		PLC_SYS_TICK_CNT :	DINT;
	END_VAR
  	RESOURCE Res0 ON PLC
    	TASK task0(INTERVAL := T#20ms,PRIORITY := 0);
    	PROGRAM instance0 WITH task0 : program0;
  	END_RESOURCE
END_CONFIGURATION

(* ---- TC_MS.ST ---- *)
FUNCTION_BLOCK T_PLC_MS_block

	VAR_OUTPUT
		T_PLC_MS :	UDINT;
	END_VAR

	VAR_EXTERNAL
		PLC_TICKS_PER_SEC :	INT;
		PLC_SYS_TICK_CNT :	DINT;
	END_VAR

	VAR
		debug :	BOOL;(*Debug-Mode ON / OFF*)
		N :	INT;(*Debug-Faktor*)
		Offset :	UDINT;(*Debug-Offset*)
		temp :	DWORD := DWORD#1;(*Debug-Offset*)
		mode :	BOOL;(*modus*)
		faktor :	UDINT;(*Systemtakt-Faktor*)
		init :	BOOL;
		v_plc_ticks_per_sec :	UDINT;
		base :	UDINT := UDINT#1000;
	END_VAR

	IF init = FALSE THEN
		v_plc_ticks_per_sec := INT_TO_UDINT(PLC_TICKS_PER_SEC);
		IF v_plc_ticks_per_sec = UDINT#1024 THEN
			faktor := UDINT#1;
			mode := FALSE;
		ELSIF v_plc_ticks_per_sec > UDINT#0 THEN
			IF v_plc_ticks_per_sec <= base THEN
				faktor := base / v_plc_ticks_per_sec;
				mode := FALSE;
			ELSE
				faktor := v_plc_ticks_per_sec / base;
				mode := TRUE;
			END_IF;
		ELSE
			faktor := UDINT#1;
		END_IF;
		init := TRUE;
	END_IF;

	IF mode THEN
		T_PLC_MS := DINT_TO_UDINT(PLC_SYS_TICK_CNT) / faktor;
	ELSE
		T_PLC_MS := DINT_TO_UDINT(PLC_SYS_TICK_CNT) * faktor;
	END_IF;

	IF debug THEN
		T_PLC_MS := (DWORD_TO_UDINT(SHL(UDINT_TO_DWORD(T_PLC_MS),N) OR SHL(temp,N)) - UDINT#1) + Offset;
	END_IF;

END_FUNCTION_BLOCK

FUNCTION_BLOCK TC_MS_Block

	VAR_OUTPUT
		TC :	DWORD;
	END_VAR

	VAR
		init :	BOOL;
		tx :	UDINT;
		last :	UDINT;
		T_PLC_MS :	T_PLC_MS_block;
	END_VAR

	T_PLC_MS();
	tx:= T_PLC_MS.T_PLC_MS;

	IF NOT init THEN
		init := TRUE;
		TC := DWORD#0;
	ELSE
		tc := UDINT_TO_DWORD(tx - last);
	END_IF;
	last := tx;

END_FUNCTION_BLOCK

PROGRAM program0

	VAR
		TC :	DWORD;
		func_block : TC_MS_Block;
	END_VAR
		func_block();
		TC := func_block.TC;

END_PROGRAM

CONFIGURATION Config0

	VAR_GLOBAL
		PLC_TICKS_PER_SEC :	INT;
		PLC_SYS_TICK_CNT :	DINT;
	END_VAR

  	RESOURCE Res0 ON PLC
    	TASK task0(INTERVAL := T#20ms,PRIORITY := 0);
    	PROGRAM instance0 WITH task0 : program0;
  	END_RESOURCE

END_CONFIGURATION

(* ---- TC_S.ST ---- *)
FUNCTION_BLOCK T_PLC_US_Block
	VAR_OUTPUT
		T_PLC_US :	UDINT;
	END_VAR

	VAR_EXTERNAL
		PLC_TICKS_PER_SEC :	INT;
		PLC_SYS_TICK_CNT :	DINT;
	END_VAR

	VAR
		debug :	BOOL;
		N :	INT;
		Offset :	UDINT;
		temp :	DWORD := DWORD#1;
		mode :	BOOL;
		faktor :	UDINT;
		init :	BOOL;
		v_plc_ticks_per_sec :	UDINT;
		base :	UDINT := UDINT#1000000;
	END_VAR

	IF init = FALSE THEN
		v_plc_ticks_per_sec := INT_TO_UDINT(PLC_TICKS_PER_SEC);
		IF v_plc_ticks_per_sec = UDINT#1024 THEN
			faktor := UDINT#1000;
			mode := FALSE;
		ELSIF v_plc_ticks_per_sec > UDINT#0 THEN
			IF v_plc_ticks_per_sec <= base THEN
				faktor := base / v_plc_ticks_per_sec;
				mode := FALSE;
			ELSE
				faktor := v_plc_ticks_per_sec / base;
				mode := TRUE;
			END_IF;
		ELSE
			faktor := UDINT#1;
		END_IF;
		init := TRUE;
	END_IF;

	IF mode THEN
		T_PLC_US := DINT_TO_UDINT(PLC_SYS_TICK_CNT) / faktor;
	ELSE
		T_PLC_US := DINT_TO_UDINT(PLC_SYS_TICK_CNT) * faktor;
	END_IF;

	IF debug THEN
		T_PLC_US := (DWORD_TO_UDINT(SHL(UDINT_TO_DWORD(T_PLC_US),N) OR SHL(temp,N)) - UDINT#1) + Offset;
	END_IF;
END_FUNCTION_BLOCK

FUNCTION_BLOCK TC_S_Block

	VAR_OUTPUT
		TC :	REAL;
	END_VAR

	VAR
		init :	BOOL;
		tx :	UDINT;
		last :	UDINT;
		T_PLC_US :	T_PLC_US_Block;
	END_VAR

	T_PLC_US();
	tx:= T_PLC_US.T_PLC_US;

	IF NOT init THEN
		init := TRUE;
		TC := 0.0;
	ELSE
		tc := UDINT_TO_REAL(tx - last) * 1.0E-6;
	END_IF;
	last := tx;

END_FUNCTION_BLOCK

PROGRAM program0

	VAR
		TC :	REAL;
		func_block : TC_S_Block;
	END_VAR
		func_block();
		TC := func_block.TC;

END_PROGRAM

CONFIGURATION Config0

	VAR_GLOBAL
		PLC_TICKS_PER_SEC :	INT;
		PLC_SYS_TICK_CNT :	DINT;
	END_VAR

	RESOURCE Res0 ON PLC
		TASK task0(INTERVAL := T#20ms,PRIORITY := 0);
		PROGRAM instance0 WITH task0 : program0;
	END_RESOURCE

END_CONFIGURATION

(* ---- TC_US.ST ---- *)
FUNCTION_BLOCK T_PLC_US_Block
	VAR_OUTPUT
		T_PLC_US :	UDINT;
	END_VAR

	VAR_EXTERNAL
		PLC_TICKS_PER_SEC :	INT;
		PLC_SYS_TICK_CNT :	DINT;
	END_VAR

	VAR
		debug :	BOOL;
		N :	INT;
		Offset :	UDINT;
		temp :	DWORD := DWORD#1;
		mode :	BOOL;
		faktor :	UDINT;
		init :	BOOL;
		v_plc_ticks_per_sec :	UDINT;
		base :	UDINT := UDINT#1000000;
	END_VAR

	IF init = FALSE THEN
		v_plc_ticks_per_sec := INT_TO_UDINT(PLC_TICKS_PER_SEC);
		IF v_plc_ticks_per_sec = UDINT#1024 THEN
			faktor := UDINT#1000;
			mode := FALSE;
		ELSIF v_plc_ticks_per_sec > UDINT#0 THEN
			IF v_plc_ticks_per_sec <= base THEN
				faktor := base / v_plc_ticks_per_sec;
				mode := FALSE;
			ELSE
				faktor := v_plc_ticks_per_sec / base;
				mode := TRUE;
			END_IF;
		ELSE
			faktor := UDINT#1;
		END_IF;
		init := TRUE;
	END_IF;

	IF mode THEN
		T_PLC_US := DINT_TO_UDINT(PLC_SYS_TICK_CNT) / faktor;
	ELSE
		T_PLC_US := DINT_TO_UDINT(PLC_SYS_TICK_CNT) * faktor;
	END_IF;

	IF debug THEN
		T_PLC_US := (DWORD_TO_UDINT(SHL(UDINT_TO_DWORD(T_PLC_US),N) OR SHL(temp,N)) - UDINT#1) + Offset;
	END_IF;
END_FUNCTION_BLOCK

FUNCTION_BLOCK TC_US_Block
	VAR_OUTPUT
		TC :	DWORD;
	END_VAR

	VAR
		init :	BOOL;
		tx :	UDINT;
		last :	UDINT;
		T_PLC_US :	T_PLC_US_Block;
	END_VAR

	T_PLC_US();
	tx:= T_PLC_US.T_PLC_US;

	IF NOT init THEN
		init := TRUE;
		TC := DWORD#0;
	ELSE
		tc := UDINT_TO_DWORD(tx - last);
	END_IF;
	last := tx;
END_FUNCTION_BLOCK

PROGRAM program0

	VAR
		TC : DWORD;
		func_block : TC_US_Block;
	END_VAR
		func_block();
		TC := func_block.TC;

END_PROGRAM

CONFIGURATION Config0
	VAR_GLOBAL
		PLC_TICKS_PER_SEC :	INT;
		PLC_SYS_TICK_CNT :	DINT;
	END_VAR

	RESOURCE Res0 ON PLC
		TASK task0(INTERVAL := T#20ms,PRIORITY := 0);
		PROGRAM instance0 WITH task0 : program0;
	END_RESOURCE
END_CONFIGURATION

(* ---- TELNET_LOG.ST ---- *)
FUNCTION_BLOCK TELNET_LOG

	VAR_INPUT
		ENABLE :	BOOL;
		OPTION :	BYTE := BYTE#2#1000_1100;
		PORT :	WORD := WORD#23;
	END_VAR

	VAR_OUTPUT
		READY :	BOOL;
	END_VAR

	VAR_IN_OUT
		IP_C :	oscat_IP_C;
		S_BUF :	oscat_NETWORK_BUFFER;
		LOG_CL :	us_LOG_CONTROL;
	END_VAR

	VAR
		TELNET_PRINT :	TELNET_PRINT;
		done :	BOOL;
		init :	BOOL;
		watchdog :	TON;
		ci :	INT;
		pi :	INT;
		pi_last :	INT;
		send :	BOOL;
	END_VAR

	IF NOT init THEN
		init := TRUE;
		IF OPTION > BYTE#0 THEN
			TELNET_PRINT.OPTION := OPTION;
		END_IF;
		IF PORT > WORD#0 THEN
			TELNET_PRINT.PORT := PORT;
		END_IF;
		WATCHDOG.PT := T#1ms;
	END_IF;

	WATCHDOG(IN:=FALSE);

	ci := LOG_CL.IDX;

	IF IP_C.C_STATE = BYTE#1 THEN
		pi := 0;
		init := FALSE;
	END_IF;

	REPEAT
		IF pi <> ci AND IP_C.C_STATE > BYTE#127 THEN
			IF pi = 0 AND LOG_CL.RING_MODE THEN pi := ci; END_IF;
			pi_last := pi;
			pi := pi + 1;
			IF pi > LOG_CL.SIZE THEN pi := 1; END_IF;
			SEND := TRUE;
		ELSE
			SEND := FALSE;
		END_IF;

		TELNET_PRINT(	IP_C := IP_C,
						S_BUF := S_BUF,
						ENABLE := ENABLE,
						SEND := SEND,
						TEXT := LOG_CL.MSG[pi],
						BACK_COLOR := DWORD_TO_BYTE(SHL(LOG_CL.MSG_OPTION[pi],8)),
						FRONT_COLOR := DWORD_TO_BYTE(LOG_CL.MSG_OPTION[pi] ));
		READY := TELNET_PRINT.READY;
		done  := TELNET_PRINT.DONE;
		IP_C  := TELNET_PRINT.IP_C;
		S_BUF := TELNET_PRINT.S_BUF;

		IF SEND AND NOT done THEN
			pi := pi_last;
		END_IF;

		WATCHDOG(IN:=TRUE);

	UNTIL (WATCHDOG.Q OR NOT done )
	END_REPEAT;

END_FUNCTION_BLOCK

(* ---- TELNET_PRINT.ST ---- *)
TYPE
  oscat_STRING250             : STRING;
END_TYPE

TYPE
  oscat_IP_FIFO128_DATA  : ARRAY [1..128] OF BYTE;
  oscat_Mailbox  : ARRAY [1..16] OF BYTE;

  oscat_IP_FIFO_DATA :
  STRUCT
	X       : oscat_IP_FIFO128_DATA; (* IP_ID FIFO Speicher          *)
	Y       : oscat_IP_FIFO128_DATA; (* IP_ID Z�hler                 *)
	ID      : BYTE;                  (* h�chste vergabene id         *)
	MAX_ID  : BYTE;                  (* maximal Anmeldungen pro ID   *)
    INIT    : BOOL;                  (* Initialisierung durchgef�hrt *)
	EMPTY   : BOOL;                  (* FIFO leer                    *)
	FULL    : BOOL;                  (* FIFO voll                    *)
	TOP     : INT;                   (* maximale anzahl in FIFO      *)
	NW      : INT;                   (* Schreibzeiger                *)
	NR      : INT;                   (* Lesezeiger                   *)
  END_STRUCT;

  oscat_IP_C:
  STRUCT
  	C_MODE:			BYTE;          		(*W Mode: TCP/UCP AKTIV/PASSIV                               *)
	C_PORT:         WORD;          		(*W Portnummer                                               *)
	C_IP:           DWORD;         		(*W IP-Adresse gepackt wwxxyyzz = www.xxx.yyy.zzz            *)
    C_STATE:        BYTE;          		(*R Verbindungsstatus ON/OFF + Flanke ON/OFF                 *)
	C_ENABLE:       BOOL;          		(*W Freigabe f�r Connect                                     *)
    R_OBSERVE:      BOOL;          		(*W Empfang ueberwachen                                      *)
    TIME_RESET:     BOOL;          		(*W Alle Timer ruecksetzen                                   *)
	ERROR:          DWORD;         		(*R vvwwxxyy (vv = CON_ERROR, ww = SEN_ERROR, xx = REC_ERROR *)
    FIFO:           oscat_IP_FIFO_DATA; (*I IP FIFO Struktur                                         *)
	MAILBOX:		oscat_Mailbox;		(*I Mailbox: Datenbereich f�r Bausteindatenaustausch         *)
  END_STRUCT;
END_TYPE

FUNCTION _BYTE_TO_INT:INT
	VAR_INPUT
		IN :	BYTE;
	END_VAR

	_BYTE_TO_INT := USINT_TO_INT(BYTE_TO_USINT(IN));
END_FUNCTION

FUNCTION_BLOCK IP_FIFO_Block

  VAR_IN_OUT
    FIFO :	oscat_IP_FIFO_DATA;
    ID :	BYTE;
    STATE :	BYTE;
  END_VAR

  VAR
    tmp :	INT;
  END_VAR

  IF NOT FIFO.INIT THEN
    FIFO.INIT		:= TRUE;
    FIFO.NW		:= 1;
    FIFO.NR		:= 1;
    FIFO.EMPTY	:= TRUE;
    FIFO.FULL		:= FALSE;
    FIFO.TOP		:= 128;
    FIFO.MAX_ID	:= BYTE#1;
  END_IF;

  IF ID = BYTE#00 THEN
    IF FIFO.ID < INT_TO_BYTE(FIFO.TOP) THEN
      ID := USINT_TO_BYTE(BYTE_TO_USINT(FIFO.ID) + USINT#1);
      FIFO.ID := ID ;

    ELSIF STATE < BYTE#200 THEN
      STATE := BYTE#255;
    RETURN;
    END_IF;
  END_IF;

  IF STATE = BYTE#1 AND NOT FIFO.FULL THEN
    tmp := _BYTE_TO_INT(ID);
    IF FIFO.Y[tmp] < FIFO.MAX_ID THEN
      FIFO.Y[tmp] := USINT_TO_BYTE(BYTE_TO_USINT(FIFO.Y[tmp]) + USINT#1);
      tmp := FIFO.NW;
      FIFO.X[tmp] := ID;
      IF FIFO.NW = FIFO.TOP THEN FIFO.NW := 1; ELSE FIFO.NW := FIFO.NW + 1; END_IF;
      FIFO.FULL := FIFO.NW = FIFO.NR;
    FIFO.EMPTY := FALSE;
      STATE := BYTE#2;
    END_IF;
  END_IF;

  IF STATE = BYTE#2 AND NOT FIFO.EMPTY THEN
    tmp := FIFO.NR;
    IF ID = FIFO.X[tmp] THEN
      STATE := BYTE#3;
    END_IF;
  END_IF;

  IF STATE = BYTE#4 AND NOT FIFO.EMPTY THEN

    tmp := FIFO.NR;
    IF ID = FIFO.X[tmp] THEN
      tmp := _BYTE_TO_INT(ID);
      FIFO.Y[tmp] := USINT_TO_BYTE(BYTE_TO_USINT(FIFO.Y[tmp]) - USINT#1);

      IF FIFO.NR = FIFO.TOP THEN FIFO.NR := 1; ELSE FIFO.NR := FIFO.NR + 1; END_IF;
      FIFO.EMPTY := FIFO.NR = FIFO.NW;
    FIFO.FULL := FALSE;
    END_IF;
    STATE := BYTE#5;
  END_IF;

END_FUNCTION_BLOCK

FUNCTION_BLOCK TELNET_PRINT_Block

	VAR_INPUT
		TEXT :	oscat_STRING250;
		ENABLE :	BOOL;
		SEND :	BOOL;
		OPTION :	BYTE;
		BACK_COLOR :	BYTE;
		FRONT_COLOR :	BYTE;
		X_POS :	BYTE;
		Y_POS :	BYTE;
		PORT :	WORD := WORD#23;
	END_VAR

	VAR_OUTPUT
		READY :	BOOL;
		DONE :	BOOL;
	END_VAR

	VAR_IN_OUT
		IP_C :	oscat_IP_C;
		S_BUF :	oscat_NETWORK_BUFFER;
	END_VAR

	VAR
		_STRING_TO_BUFFER :	_STRING_TO_BUFFER_NW;
		last_fc :	BYTE;
		state :	INT;
		x :	INT := -1;
		ip_state :	BYTE;
		ip_id :	BYTE;
		IP_FIFO :	IP_FIFO_Block;
		s_buf_size :	UINT := uint#4096;
		init :	BOOL;
		b0_screen_clear :	BOOL;
		b1_autowrap :	BOOL;
		b2_color :	BOOL;
		b3_cr_lr :	BOOL;
		b7_no_flush :	BOOL;
	END_VAR

	READY := IP_C.C_STATE > BYTE#127;
	DONE := FALSE;

	CASE state OF

	00:
		IF ENABLE THEN
			state := 10;
			ip_state := BYTE#1;
		END_IF;

	10:
		IF ip_state = BYTE#3 THEN

			IP_C.C_PORT := PORT;
			IP_C.C_IP := DWORD#00;
			IP_C.C_MODE := BYTE#4;
			IP_C.TIME_RESET := TRUE;
			IP_C.C_ENABLE := TRUE;
			IP_C.R_OBSERVE := FALSE;
			state := 20;
		END_IF;

	20:	IF IP_C.ERROR > DWORD#0 THEN
			IP_C.TIME_RESET := TRUE;
		END_IF;
		IF S_BUF.SIZE = UINT#0 THEN
			IF NOT ENABLE THEN
				ip_state := BYTE#4;
				IP_C.C_ENABLE := FALSE;
				state := 0;
			END_IF;
			IF IP_C.C_STATE = BYTE#1 THEN
				init := FALSE;
			ELSIF READY THEN
				IF IP_C.C_STATE = BYTE#254 AND NOT INIT THEN
					init := TRUE;
					b0_screen_clear := (OPTION AND BYTE#2#0000_0001) > BYTE#0;
					b1_autowrap := (OPTION AND BYTE#2#0000_0010) > BYTE#0;
					b2_color := (OPTION AND BYTE#2#0000_0100) > BYTE#0;
					b3_cr_lr := (OPTION AND BYTE#2#0000_1000) > BYTE#0;
					b7_no_flush := (OPTION AND BYTE#2#1000_0000) > BYTE#0;

					last_fc := NOT FRONT_COLOR;
					x := 0;

					S_BUF.BUFFER[x] := BYTE#16#1B;
					x := x +1;
					S_BUF.BUFFER[x] := BYTE#16#5B;
					x := x +1;
					S_BUF.BUFFER[x] := BYTE#16#3F;
					x := x +1;
					S_BUF.BUFFER[x] := BYTE#16#37; (
					x := x +1;
					S_BUF.BUFFER[x] := SEL(b1_autowrap, BYTE#16#6C, BYTE#16#68 );

					IF b0_screen_clear THEN
						IF b2_color THEN
							x := x +1;
							S_BUF.BUFFER[x] := BYTE#16#1B;
							x := x +1;
							S_BUF.BUFFER[x] := BYTE#16#5B;
							x := x +1;
							S_BUF.BUFFER[x] := BYTE#16#30;
							x := x +1;
							S_BUF.BUFFER[x] := BYTE#16#3B;
							x := x +1;
							S_BUF.BUFFER[x] := BYTE#16#33;
							x := x +1;
							S_BUF.BUFFER[x] := (FRONT_COLOR AND BYTE#2#00000111) OR BYTE#16#30;
							x := x +1;
							S_BUF.BUFFER[x] := BYTE#16#3B;
							x := x +1;
							S_BUF.BUFFER[x] := BYTE#16#34;
							x := x +1;
							S_BUF.BUFFER[x] := (BACK_COLOR AND BYTE#2#00000111) OR BYTE#16#30;
							x := x +1;
							S_BUF.BUFFER[x] := BYTE#16#6D;
						END_IF;
						x := x +1;
						S_BUF.BUFFER[x] := BYTE#16#1B;
						x := x +1;
						S_BUF.BUFFER[x] := BYTE#16#5B;
						x := x +1;
						S_BUF.BUFFER[x] := BYTE#16#32;
						x := x +1;
						S_BUF.BUFFER[x] := BYTE#16#4A;
					ELSE
						x := x +1;
						S_BUF.BUFFER[x] := BYTE#16#0A;
					END_IF;
				END_IF;

				IF (INT_TO_UINT(x + LEN(TEXT) + 21) > s_buf_size) OR (x >= 0 AND NOT SEND) THEN
					S_BUF.SIZE := INT_TO_UINT(x + 1);
					x := -1;
				ELSIF SEND THEN

					IF b2_color AND FRONT_COLOR <> last_FC THEN
						x := x + 1;
						S_BUF.BUFFER[x] := BYTE#16#1B;
						x := x + 1;
						S_BUF.BUFFER[x] := BYTE#16#5B;
						IF ((FRONT_COLOR AND BYTE#2#0001_1000) XOR (last_FC AND BYTE#2#0001_1000)) <> BYTE#00 OR TRUE THEN
							x := x + 1;
							S_BUF.BUFFER[x] := BYTE#16#30;
							x := x + 1;
							S_BUF.BUFFER[x] := BYTE#16#3B;
							IF (FRONT_COLOR AND BYTE#2#00001000) = BYTE#0 THEN
								x := x + 1;
								S_BUF.BUFFER[x] := BYTE#16#31;
								x := x + 1;
								S_BUF.BUFFER[x] := BYTE#16#3B;
							END_IF;
							IF (FRONT_COLOR AND BYTE#2#00010000) > BYTE#0 THEN
								x := x + 1;
								S_BUF.BUFFER[x] := BYTE#16#35;
								x := x + 1;
								S_BUF.BUFFER[x] := BYTE#16#3B;
							END_IF;
						END_IF;
						x := x + 1;
						S_BUF.BUFFER[x] := BYTE#16#33;
						x := x + 1;
						S_BUF.BUFFER[x] := (FRONT_COLOR AND BYTE#2#00000111) OR BYTE#16#30;
						x := x + 1;
						S_BUF.BUFFER[x] := BYTE#16#6D;
						last_FC := FRONT_COLOR;
					END_IF;

					IF X_POS > BYTE#0 AND Y_POS > BYTE#0 THEN
						x := x + 1;
						S_BUF.BUFFER[x] := BYTE#16#1B;
						x := x + 1;
						S_BUF.BUFFER[x] := BYTE#16#5B;
						x := x + 1;
						S_BUF.BUFFER[x] := SHR(INT_TO_BCDC(BYTE_TO_INT(Y_POS)),4) OR BYTE#16#30;
						x := x + 1;
						S_BUF.BUFFER[x] := (INT_TO_BCDC(BYTE_TO_INT(Y_POS)) AND BYTE#16#0F) OR BYTE#16#30;
						x := x + 1;
						S_BUF.BUFFER[x] := BYTE#16#3B;
						x := x + 1;
						S_BUF.BUFFER[x] := SHR(INT_TO_BCDC(BYTE_TO_INT(X_POS)),4) OR BYTE#16#30;
						x := x + 1;
						S_BUF.BUFFER[x] := (INT_TO_BCDC(BYTE_TO_INT(X_POS)) AND BYTE#16#0F) OR BYTE#16#30;
						x := x + 1;
						S_BUF.BUFFER[x] := BYTE#16#48;
					END_IF;

					IF LEN(TEXT) > 0 THEN
						_STRING_TO_BUFFER(str:=TEXT,pos:=x + 1,size:=s_buf_size,pt:=S_BUF.BUFFER);
						S_BUF.BUFFER:=_STRING_TO_BUFFER.pt;
						x := x + LEN(TEXT);
					END_IF;

					IF b3_cr_lr THEN
						x := x + 1;
						S_BUF.BUFFER[x] := BYTE#16#0D;
						x := x + 1;
						S_BUF.BUFFER[x] := BYTE#16#0A;
					END_IF;

					DONE := TRUE;

					IF b7_no_flush THEN
						S_BUF.SIZE := INT_TO_UINT(x + 1);
						x := -1;
					END_IF;
				END_IF;
			END_IF;
		END_IF;
	END_CASE;

	IP_FIFO(FIFO:=IP_C.FIFO,STATE:=IP_STATE,ID:=IP_ID);
	IP_C.FIFO:=IP_FIFO.FIFO;
	IP_STATE := IP_FIFO.STATE;
	IP_ID:=IP_FIFO.ID;

	READY := IP_C.C_STATE > BYTE#127;
	DONE := FALSE;

	CASE state OF

	00:
		IF ENABLE THEN
			state := 10;
			IP_STATE := BYTE#1;
		END_IF;

	10:
		IF IP_STATE = BYTE#3 THEN

			IP_C.C_PORT     := WORD#23;
			IP_C.C_IP       := DWORD#00;
			IP_C.C_MODE     := BYTE#4;
			IP_C.TIME_RESET := TRUE;
			IP_C.C_ENABLE   := TRUE;
			IP_C.R_OBSERVE  := FALSE;
			state := 20;
		END_IF;

	20: IF IP_C.ERROR > DWORD#0 THEN
			IP_C.TIME_RESET := TRUE;
		END_IF;
		IF S_BUF.SIZE = UINT#0 THEN
			IF NOT ENABLE THEN
				IP_STATE := BYTE#4;
				IP_C.C_ENABLE := FALSE;
				state := 0;
			END_IF;
			IF IP_C.C_STATE = BYTE#1  THEN
				INIT := FALSE;
			ELSIF READY THEN
				IF IP_C.C_STATE = BYTE#254 AND NOT INIT THEN
					INIT := TRUE;
					last_FC := NOT FRONT_COLOR;

					_STRING_TO_BUFFER(str:='#[?7h#[0;3#;4#m#[2J',pos:=0,size:=S_BUF_SIZE,pt:=S_BUF.BUFFER);
					S_BUF.BUFFER:=_STRING_TO_BUFFER.pt;

					S_BUF.BUFFER[0] := BYTE#16#1B;
					IF (OPTION AND BYTE#2#0000_0010) > BYTE#0 THEN
						S_BUF.BUFFER[4] := BYTE#16#6C;
					END_IF;
					x := 4;
					IF (OPTION AND BYTE#2#0000_0001) > BYTE#0 THEN

						S_BUF.BUFFER[05] := BYTE#16#1B;
						S_BUF.BUFFER[10] := (FRONT_COLOR AND BYTE#2#00000111) OR BYTE#16#30;
						S_BUF.BUFFER[13] := (BACK_COLOR AND BYTE#2#00000111) OR BYTE#16#30;
						S_BUF.BUFFER[15] := BYTE#16#1B;
						x := 18;
					ELSE
						x := x + 1;
						S_BUF.BUFFER[x] := BYTE#16#0A;
					END_IF;
				END_IF;

				IF (INT_TO_UINT(x + LEN(TEXT) + 21) > S_BUF_SIZE) OR (x >= 0 AND NOT SEND) THEN
					S_BUF.SIZE := INT_TO_UINT(x + 1);
					x := -1;
				ELSIF SEND THEN

					IF (OPTION AND BYTE#2#0000_0100) > BYTE#0 AND FRONT_COLOR <> last_FC THEN
						x := x + 1;
						S_BUF.BUFFER[x] := BYTE#16#1B;
						x := x + 1;
						S_BUF.BUFFER[x] := BYTE#16#5B;
						IF ((FRONT_COLOR AND BYTE#2#0001_1000) XOR (last_FC AND BYTE#2#0001_1000)) <> BYTE#00 OR TRUE THEN
							x := x + 1;
							S_BUF.BUFFER[x] := BYTE#16#30;
							x := x + 1;
							S_BUF.BUFFER[x] := BYTE#16#3B;
							IF (FRONT_COLOR AND BYTE#2#00001000) = BYTE#0 THEN
								x := x + 1;
								S_BUF.BUFFER[x] := BYTE#16#31;
								x := x + 1;
								S_BUF.BUFFER[x] := BYTE#16#3B;
							END_IF;
							IF (FRONT_COLOR AND BYTE#2#00010000) > BYTE#0 THEN
								x := x + 1;
								S_BUF.BUFFER[x] := BYTE#16#35;
								x := x + 1;
								S_BUF.BUFFER[x] := BYTE#16#3B;
							END_IF;
						END_IF;
						x := x + 1;
						S_BUF.BUFFER[x] := BYTE#16#33;
						x := x + 1;
						S_BUF.BUFFER[x] := (FRONT_COLOR AND BYTE#2#00000111) OR BYTE#16#30;
						x := x + 1;
						S_BUF.BUFFER[x] := BYTE#16#6D;
						last_FC := FRONT_COLOR;
					END_IF;

					IF X_POS > BYTE#0 AND Y_POS > BYTE#0 THEN
						x := x + 1;
						S_BUF.BUFFER[x] := BYTE#16#1B;
						x := x + 1;
						S_BUF.BUFFER[x] := BYTE#16#5B;
						x := x + 1;
						S_BUF.BUFFER[x] := SHR_BYTE(INT_TO_BCDC(_BYTE_TO_INT(Y_POS)),4) OR BYTE#16#30;
						x := x + 1;
						S_BUF.BUFFER[x] := (INT_TO_BCDC(_BYTE_TO_INT(Y_POS)) AND BYTE#16#0F) OR BYTE#16#30;
						x := x + INT#1;
						S_BUF.BUFFER[x] := BYTE#16#3B;
						x := x + 1;
						S_BUF.BUFFER[x] := SHR_BYTE(INT_TO_BCDC(_BYTE_TO_INT(X_POS)),4) OR BYTE#16#30;
						x := x + 1;
						S_BUF.BUFFER[x] := (INT_TO_BCDC(_BYTE_TO_INT(X_POS)) AND BYTE#16#0F) OR BYTE#16#30;
						x := x + 1;
						S_BUF.BUFFER[x] := BYTE#16#48;
					END_IF;

					IF LEN(TEXT) > 0 THEN

						_STRING_TO_BUFFER(str:=TEXT,pos:=x + 1,size:=S_BUF_SIZE,pt:=S_BUF.BUFFER);
						S_BUF.BUFFER:=_STRING_TO_BUFFER.pt;
						x := x + LEN(TEXT);
					END_IF;

					IF (OPTION AND BYTE#2#0000_1000) > BYTE#0 THEN
						x := x + 1;
						S_BUF.BUFFER[x] := BYTE#16#0D;
						x := x + 1;
						S_BUF.BUFFER[x] := BYTE#16#0A;
					END_IF;

					DONE := TRUE;

					IF (OPTION AND BYTE#2#1000_0000) = BYTE#0 THEN
						S_BUF.SIZE := INT_TO_UINT(x + 1);
						x := -1;
					END_IF;
				END_IF;
			END_IF;
		END_IF;
	END_CASE;

	IP_FIFO(FIFO:=IP_C.FIFO,STATE:=IP_STATE,ID:=IP_ID);
	IP_C.FIFO:=IP_FIFO.FIFO;
	IP_STATE := IP_FIFO.STATE;
	IP_ID:=IP_FIFO.ID;

END_FUNCTION_BLOCK

PROGRAM program0
	VAR
		TEXT :	oscat_STRING250;
		ENABLE :	BOOL;
		SEND :	BOOL;
		OPTION :	BYTE;
		BACK_COLOR :	BYTE;
		FRONT_COLOR :	BYTE;
		X_POS :	BYTE;
		Y_POS :	BYTE;
		PORT :	WORD := WORD#23;
		IP_C :	oscat_IP_C;
		S_BUF :	oscat_NETWORK_BUFFER;
		READY :	BOOL;
		DONE :	BOOL;

		func_block : TELNET_PRINT_Block;
	END_VAR
	func_block.TEXT := TEXT;
	func_block.ENABLE := ENABLE;
	func_block.SEND := SEND;
	func_block.OPTION := OPTION;
	func_block.BACK_COLOR := BACK_COLOR;
	func_block.FRONT_COLOR := FRONT_COLOR;
	func_block.X_POS := X_POS;
	func_block.Y_POS := Y_POS;
	func_block.PORT := PORT;
	func_block.IP_C := IP_C;
	func_block.S_BUF := S_BUF;

	func_block();
	IP_C  := func_block.IP_C;
	S_BUF  := func_block.S_BUF;
	READY  := func_block.READY;
	DONE  := func_block.DONE;
END_PROGRAM

CONFIGURATION Config0
	RESOURCE Res0 ON PLC
		TASK task0(INTERVAL := T#20ms,PRIORITY := 0);
		PROGRAM instance0 WITH task0 : program0;
	END_RESOURCE
END_CONFIGURATION
